IF GVL_HMI.rRobotManualSpeedPercent < REAL#0.1 THEN
	GVL_HMI.rRobotManualSpeedPercent := REAL#0.1;
ELSIF GVL_HMI.rRobotManualSpeedPercent > REAL#100.0 THEN
	GVL_HMI.rRobotManualSpeedPercent := REAL#100.0;
END_IF;
IF (GVL_HMI.lrRobotManualStep <> 0.1)
AND (GVL_HMI.lrRobotManualStep <> 1.0)
AND (GVL_HMI.lrRobotManualStep <> 10.0)
AND (GVL_HMI.lrRobotManualStep <> 100.0) THEN
	GVL_HMI.lrRobotManualStep := 1.0;
END_IF;

IF NOT xHmiConnectionAlive THEN
	FOR uiMachine := 1 TO 3 DO
		GVL_HMI.astAxisHmiCommand[uiMachine].xJogPositive := FALSE;
		GVL_HMI.astAxisHmiCommand[uiMachine].xJogNegative := FALSE;
		GVL_HMI.astAxisHmiCommand[uiMachine].xHome := FALSE;
		GVL_HMI.astAxisHmiCommand[uiMachine].xMoveAbsolute := FALSE;
		GVL_HMI.astAxisHmiCommand[uiMachine].xMoveRelative := FALSE;
	END_FOR;
	FOR uiMagazine := UINT#1 TO UINT#2 DO
		GVL_HMI.astMagazineCommand[uiMagazine].xStop := FALSE;
	END_FOR;
	GVL_HMI.xRobotManualExecute := FALSE;
END_IF;

// Глобальные команды ячейки поступают через единый интерфейс HMI.
GVL_CELL_CONTROL.xEnable := GVL_HMI.xCellEnable;
GVL_CELL_CONTROL.xDisable := GVL_HMI.xCellDisable;
GVL_CELL_CONTROL.xStart := GVL_HMI.xCellStart;
GVL_CELL_CONTROL.xStop := GVL_HMI.xCellStop;
// Необработанный общий импульс передаётся всем владельцам аварий.
// Каждый функциональный блок самостоятельно проверяет возможность сброса.
GVL_CELL_CONTROL.xReset := GVL_HMI.xCellReset;
// Режим хранит PLC. Новая транзакция применяется в RunSafety после чтения
// актуальных входов безопасности; PublishHmi не пишет в буфер запроса.
GVL_ALARM.Command.xResetWarnings := GVL_HMI.xAlarmResetWarnings;

// Режим инъекции ошибок включается отдельным переключателем страницы CELL_SETTINGS.
GVL_CELL_SETTINGS.xErrorSimulationEnabled := GVL_HMI.xErrorSimulationEnable
	AND (GVL_CELL_SETTINGS.eTestEnvironment <> E_CELL_TEST_ENVIRONMENT.NORMAL);

// Ползунок меняет только запрошенное значение. Отдельный FB применяет его к
// таймерам и Dynamic Limits безопасной транзакцией перед следующим тестом.
GVL_CELL_SETTINGS.xSimulationAccelerationChangeAllowed :=
	xHmiConnectionAlive
	AND NOT GVL_CELL_CONTROL.xGlobalError;

IF GVL_CELL_SETTINGS.xSimulationAccelerationChangeAllowed THEN
	GVL_CELL_SETTINGS.xSimulationAccelerationEnable := GVL_HMI.xSimulationAccelerationEnable;
	GVL_CELL_SETTINGS.uiSimulationTimeFactor := GVL_HMI.uiSimulationTimeFactor;
	IF GVL_CELL_SETTINGS.uiSimulationTimeFactor < UINT#1 THEN
		GVL_CELL_SETTINGS.uiSimulationTimeFactor := UINT#1;
	ELSIF GVL_CELL_SETTINGS.uiSimulationTimeFactor > UINT#100 THEN
		GVL_CELL_SETTINGS.uiSimulationTimeFactor := UINT#100;
	END_IF;
ELSE
	// При потере разрешения сохраняем последнее принятое требование.
	GVL_HMI.xSimulationAccelerationEnable := GVL_CELL_SETTINGS.xSimulationAccelerationActive;
	GVL_HMI.uiSimulationTimeFactor := GVL_CELL_SETTINGS.uiSimulationTimeFactor;
END_IF;

// Общие технологические TIMEOUT и допуски HOME принимаются только при полностью
// остановленной ячейке. Координатами HOME_SAFETY владеет редактор точек ниже.
GVL_CELL_SETTINGS.xCellSettingsChangeAllowed :=
	xHmiConnectionAlive
	AND NOT GVL_CELL_MANAGER.Status.xRunning
	AND NOT GVL_HMI.xModbusMode
	AND NOT GVL_CELL_CONTROL.xGlobalError
	AND NOT GVL_AXIS.arrAxis[1].Status.xMotionBusy
	AND NOT GVL_AXIS.arrAxis[2].Status.xMotionBusy
	AND NOT GVL_AXIS.arrAxis[3].Status.xMotionBusy
	AND NOT GVL_AXIS_GROUP.AxisGroup.Command.xMoveDirect
	AND NOT GVL_AXIS_GROUP.AxisGroup.Command.xMoveLinear
	AND NOT xPowerTransitionActive
	AND NOT SIMULATION_DYNAMICS.xBusy
	AND NOT GVL_ROBOT.Status.xBusy;

GVL_CELL_SETTINGS.xIoFilterSettingsChangeAllowed := xHmiConnectionAlive
	AND GVL_CELL_CONTROL.xManual
	AND NOT GVL_CELL_MANAGER.Status.xRunning
	AND NOT GVL_ROBOT.Status.xBusy AND NOT xMotionBusy
	AND NOT xPowerTransitionActive AND NOT SIMULATION_DYNAMICS.xBusy
	AND NOT GVL_MACHINE.Status[1].xBusy AND NOT GVL_MACHINE.Status[1].xProcessing
	AND NOT GVL_MACHINE.Status[2].xBusy AND NOT GVL_MACHINE.Status[2].xProcessing
	AND NOT GVL_MACHINE.Status[3].xBusy AND NOT GVL_MACHINE.Status[3].xProcessing
	AND NOT GVL_TWO_PALLET.astStatus[1].xBusy AND NOT GVL_TWO_PALLET.astStatus[2].xBusy
	AND NOT GVL_TWO_PALLET.astInput[1].xPowered AND NOT GVL_TWO_PALLET.astInput[2].xPowered;

// Independent requested value; publication cannot overwrite an incoming write.
xCellSettingRejected := FALSE;
udiCellSettingSnapshot := GVL_HMI.udiCellSettingCommandSeq;
IF (udiCellSettingSnapshot <> UDINT#0)
AND (udiCellSettingSnapshot <> GVL_HMI.udiCellSettingAckSeq) THEN
	GVL_HMI.uiCellSettingResult := UINT#3;
	IF NOT IsHmiCommandFresh(udiIssuedAtMs := GVL_HMI.udiCellSettingIssuedAtMs) THEN
		GVL_HMI.uiCellSettingResult := UINT#4; // Expired: never apply later
	ELSIF ((((GVL_HMI.uiCellSettingIndex = UINT#37) OR (GVL_HMI.uiCellSettingIndex = UINT#38) OR (GVL_HMI.uiCellSettingIndex = UINT#39))
		AND NOT GVL_CELL_SETTINGS.xIoFilterSettingsChangeAllowed)
		OR (((GVL_HMI.uiCellSettingIndex <> UINT#37) AND (GVL_HMI.uiCellSettingIndex <> UINT#38) AND (GVL_HMI.uiCellSettingIndex <> UINT#39))
			AND NOT GVL_CELL_SETTINGS.xCellSettingsChangeAllowed))
	OR (((GVL_HMI.uiCellSettingIndex = UINT#4)
		OR (GVL_HMI.uiCellSettingIndex = UINT#25)
		OR (GVL_HMI.uiCellSettingIndex = UINT#29))
		AND xPointCheckActive)
	OR ((GVL_HMI.uiCellSettingIndex = UINT#28) AND xMobileMotionLeaseActive) THEN
		GVL_HMI.uiCellSettingResult := UINT#2;
	ELSE
		CASE GVL_HMI.uiCellSettingIndex OF
			UINT#1:
				IF (GVL_HMI.lrCellSettingRequest >= 0.1) AND (GVL_HMI.lrCellSettingRequest <= 1000.0) THEN
					GVL_CELL_SETTINGS.lrSafetyHomeToleranceX := GVL_HMI.lrCellSettingRequest;
					GVL_HMI.uiCellSettingResult := UINT#1;
				END_IF;
			UINT#2:
				IF (GVL_HMI.lrCellSettingRequest >= 0.1) AND (GVL_HMI.lrCellSettingRequest <= 1000.0) THEN
					GVL_CELL_SETTINGS.lrSafetyHomeToleranceY := GVL_HMI.lrCellSettingRequest;
					GVL_HMI.uiCellSettingResult := UINT#1;
				END_IF;
			UINT#3:
				IF (GVL_HMI.lrCellSettingRequest >= 0.1) AND (GVL_HMI.lrCellSettingRequest <= 1000.0) THEN
					GVL_CELL_SETTINGS.lrSafetyHomeToleranceZ := GVL_HMI.lrCellSettingRequest;
					GVL_HMI.uiCellSettingResult := UINT#1;
				END_IF;
			UINT#4:
				IF (GVL_HMI.lrCellSettingRequest >= 0.1) AND (GVL_HMI.lrCellSettingRequest <= 100.0) THEN
					GVL_CELL_SETTINGS.rPointCheckSpeedPercent := LREAL_TO_REAL(GVL_HMI.lrCellSettingRequest);
					GVL_HMI.uiCellSettingResult := UINT#1;
				END_IF;
			UINT#5:
				IF (GVL_HMI.lrCellSettingRequest >= 1000.0) AND (GVL_HMI.lrCellSettingRequest <= 600000.0) THEN
					GVL_CELL_SETTINGS.stMachineTimeouts.tRobotMove := UDINT_TO_TIME(LREAL_TO_UDINT(GVL_HMI.lrCellSettingRequest));
					GVL_HMI.uiCellSettingResult := UINT#1;
				END_IF;
			UINT#6:
				IF (GVL_HMI.lrCellSettingRequest >= 1000.0) AND (GVL_HMI.lrCellSettingRequest <= 600000.0) THEN
					GVL_CELL_SETTINGS.stMachineTimeouts.tRobotAction := UDINT_TO_TIME(LREAL_TO_UDINT(GVL_HMI.lrCellSettingRequest));
					GVL_HMI.uiCellSettingResult := UINT#1;
				END_IF;
			UINT#7:
				IF (GVL_HMI.lrCellSettingRequest >= 1000.0) AND (GVL_HMI.lrCellSettingRequest <= 600000.0) THEN
					GVL_CELL_SETTINGS.stMachineTimeouts.tRobotRelease := UDINT_TO_TIME(LREAL_TO_UDINT(GVL_HMI.lrCellSettingRequest));
					GVL_HMI.uiCellSettingResult := UINT#1;
				END_IF;
			UINT#8:
				IF (GVL_HMI.lrCellSettingRequest >= 1000.0) AND (GVL_HMI.lrCellSettingRequest <= 600000.0) THEN
					GVL_CELL_SETTINGS.stMachineTimeouts.tDoorOpen := UDINT_TO_TIME(LREAL_TO_UDINT(GVL_HMI.lrCellSettingRequest));
					GVL_HMI.uiCellSettingResult := UINT#1;
				END_IF;
			UINT#9:
				IF (GVL_HMI.lrCellSettingRequest >= 1000.0) AND (GVL_HMI.lrCellSettingRequest <= 600000.0) THEN
					GVL_CELL_SETTINGS.stMachineTimeouts.tDoorClose := UDINT_TO_TIME(LREAL_TO_UDINT(GVL_HMI.lrCellSettingRequest));
					GVL_HMI.uiCellSettingResult := UINT#1;
				END_IF;
			UINT#10:
				IF (GVL_HMI.lrCellSettingRequest >= 1000.0) AND (GVL_HMI.lrCellSettingRequest <= 600000.0) THEN
					GVL_CELL_SETTINGS.stMachineTimeouts.tHatchUnlock := UDINT_TO_TIME(LREAL_TO_UDINT(GVL_HMI.lrCellSettingRequest));
					GVL_HMI.uiCellSettingResult := UINT#1;
				END_IF;
			UINT#11:
				IF (GVL_HMI.lrCellSettingRequest >= 1000.0) AND (GVL_HMI.lrCellSettingRequest <= 600000.0) THEN
					GVL_CELL_SETTINGS.stMachineTimeouts.tChuckOpen := UDINT_TO_TIME(LREAL_TO_UDINT(GVL_HMI.lrCellSettingRequest));
					GVL_HMI.uiCellSettingResult := UINT#1;
				END_IF;
			UINT#12:
				IF (GVL_HMI.lrCellSettingRequest >= 1000.0) AND (GVL_HMI.lrCellSettingRequest <= 600000.0) THEN
					GVL_CELL_SETTINGS.stMachineTimeouts.tChuckClose := UDINT_TO_TIME(LREAL_TO_UDINT(GVL_HMI.lrCellSettingRequest));
					GVL_HMI.uiCellSettingResult := UINT#1;
				END_IF;
			UINT#13:
				IF (GVL_HMI.lrCellSettingRequest >= 1000.0) AND (GVL_HMI.lrCellSettingRequest <= 600000.0) THEN
					GVL_CELL_SETTINGS.stMachineTimeouts.tCycleStart := UDINT_TO_TIME(LREAL_TO_UDINT(GVL_HMI.lrCellSettingRequest));
					GVL_HMI.uiCellSettingResult := UINT#1;
				END_IF;
			UINT#14:
				IF (GVL_HMI.lrCellSettingRequest >= 1000.0) AND (GVL_HMI.lrCellSettingRequest <= 600000.0) THEN
					GVL_CELL_SETTINGS.stAxisTimeouts.tPowerTimeout := UDINT_TO_TIME(LREAL_TO_UDINT(GVL_HMI.lrCellSettingRequest));
					GVL_HMI.uiCellSettingResult := UINT#1;
				END_IF;
			UINT#15:
				IF (GVL_HMI.lrCellSettingRequest >= 1000.0) AND (GVL_HMI.lrCellSettingRequest <= 600000.0) THEN
					GVL_CELL_SETTINGS.stAxisTimeouts.tResetTimeout := UDINT_TO_TIME(LREAL_TO_UDINT(GVL_HMI.lrCellSettingRequest));
					GVL_HMI.uiCellSettingResult := UINT#1;
				END_IF;
			UINT#16:
				IF (GVL_HMI.lrCellSettingRequest >= 1000.0) AND (GVL_HMI.lrCellSettingRequest <= 600000.0) THEN
					GVL_CELL_SETTINGS.stAxisTimeouts.tStopTimeout := UDINT_TO_TIME(LREAL_TO_UDINT(GVL_HMI.lrCellSettingRequest));
					GVL_HMI.uiCellSettingResult := UINT#1;
				END_IF;
			UINT#17:
				IF (GVL_HMI.lrCellSettingRequest >= 1000.0) AND (GVL_HMI.lrCellSettingRequest <= 600000.0) THEN
					GVL_CELL_SETTINGS.stAxisTimeouts.tHomeTimeout := UDINT_TO_TIME(LREAL_TO_UDINT(GVL_HMI.lrCellSettingRequest));
					GVL_HMI.uiCellSettingResult := UINT#1;
				END_IF;
			UINT#18:
				IF (GVL_HMI.lrCellSettingRequest >= 1000.0) AND (GVL_HMI.lrCellSettingRequest <= 600000.0) THEN
					GVL_CELL_SETTINGS.stAxisTimeouts.tMoveTimeout := UDINT_TO_TIME(LREAL_TO_UDINT(GVL_HMI.lrCellSettingRequest));
					GVL_HMI.uiCellSettingResult := UINT#1;
				END_IF;
			UINT#19:
				IF (GVL_HMI.lrCellSettingRequest >= 1000.0) AND (GVL_HMI.lrCellSettingRequest <= 600000.0) THEN
					GVL_CELL_SETTINGS.stAxisGroupTimeouts.tPowerTimeout := UDINT_TO_TIME(LREAL_TO_UDINT(GVL_HMI.lrCellSettingRequest));
					GVL_HMI.uiCellSettingResult := UINT#1;
				END_IF;
			UINT#20:
				IF (GVL_HMI.lrCellSettingRequest >= 1000.0) AND (GVL_HMI.lrCellSettingRequest <= 600000.0) THEN
					GVL_CELL_SETTINGS.stAxisGroupTimeouts.tGroupTimeout := UDINT_TO_TIME(LREAL_TO_UDINT(GVL_HMI.lrCellSettingRequest));
					GVL_HMI.uiCellSettingResult := UINT#1;
				END_IF;
			UINT#21:
				IF (GVL_HMI.lrCellSettingRequest >= 1000.0) AND (GVL_HMI.lrCellSettingRequest <= 600000.0) THEN
					GVL_CELL_SETTINGS.stAxisGroupTimeouts.tStopTimeout := UDINT_TO_TIME(LREAL_TO_UDINT(GVL_HMI.lrCellSettingRequest));
					GVL_HMI.uiCellSettingResult := UINT#1;
				END_IF;
			UINT#22:
				IF (GVL_HMI.lrCellSettingRequest >= 1000.0) AND (GVL_HMI.lrCellSettingRequest <= 600000.0) THEN
					GVL_CELL_SETTINGS.stAxisGroupTimeouts.tHaltTimeout := UDINT_TO_TIME(LREAL_TO_UDINT(GVL_HMI.lrCellSettingRequest));
					GVL_HMI.uiCellSettingResult := UINT#1;
				END_IF;
			UINT#23:
				IF (GVL_HMI.lrCellSettingRequest >= 1000.0) AND (GVL_HMI.lrCellSettingRequest <= 600000.0) THEN
					GVL_CELL_SETTINGS.stAxisGroupTimeouts.tHomeTimeout := UDINT_TO_TIME(LREAL_TO_UDINT(GVL_HMI.lrCellSettingRequest));
					GVL_HMI.uiCellSettingResult := UINT#1;
				END_IF;
			UINT#24:
				IF (GVL_HMI.lrCellSettingRequest >= 1000.0) AND (GVL_HMI.lrCellSettingRequest <= 600000.0) THEN
					GVL_CELL_SETTINGS.stAxisGroupTimeouts.tMoveTimeout := UDINT_TO_TIME(LREAL_TO_UDINT(GVL_HMI.lrCellSettingRequest));
					GVL_HMI.uiCellSettingResult := UINT#1;
				END_IF;
			UINT#25:
				IF (GVL_HMI.lrCellSettingRequest >= 500.0) AND (GVL_HMI.lrCellSettingRequest <= 60000.0) THEN
					GVL_CELL_SETTINGS.tPointCheckStartTimeout := UDINT_TO_TIME(LREAL_TO_UDINT(GVL_HMI.lrCellSettingRequest));
					GVL_HMI.uiCellSettingResult := UINT#1;
				END_IF;
			UINT#26:
				IF (GVL_HMI.lrCellSettingRequest >= 1000.0) AND (GVL_HMI.lrCellSettingRequest <= 600000.0) THEN
					GVL_CELL_SETTINGS.tSimulationDynamicsTimeout := UDINT_TO_TIME(LREAL_TO_UDINT(GVL_HMI.lrCellSettingRequest));
					GVL_HMI.uiCellSettingResult := UINT#1;
				END_IF;
			UINT#27:
				IF (GVL_HMI.lrCellSettingRequest >= 500.0) AND (GVL_HMI.lrCellSettingRequest <= 30000.0) THEN
					GVL_CELL_SETTINGS.tHmiWatchdogTimeout := UDINT_TO_TIME(LREAL_TO_UDINT(GVL_HMI.lrCellSettingRequest));
					GVL_HMI.uiCellSettingResult := UINT#1;
				END_IF;
			UINT#28:
				IF (GVL_HMI.lrCellSettingRequest >= 500.0) AND (GVL_HMI.lrCellSettingRequest <= 30000.0) THEN
					GVL_CELL_SETTINGS.tMobileMotionWatchdogTimeout := UDINT_TO_TIME(LREAL_TO_UDINT(GVL_HMI.lrCellSettingRequest));
					GVL_HMI.uiCellSettingResult := UINT#1;
				END_IF;
			UINT#29:
				IF (GVL_HMI.lrCellSettingRequest >= 500.0) AND (GVL_HMI.lrCellSettingRequest <= 30000.0) THEN
					GVL_CELL_SETTINGS.tPointCheckWatchdogTimeout := UDINT_TO_TIME(LREAL_TO_UDINT(GVL_HMI.lrCellSettingRequest));
					GVL_HMI.uiCellSettingResult := UINT#1;
				END_IF;
			UINT#30:
				IF (GVL_HMI.lrCellSettingRequest >= 1000.0) AND (GVL_HMI.lrCellSettingRequest <= 30000.0) THEN
					GVL_CELL_SETTINGS.tHmiCommandFreshnessTimeout := UDINT_TO_TIME(LREAL_TO_UDINT(GVL_HMI.lrCellSettingRequest));
					GVL_HMI.uiCellSettingResult := UINT#1;
				END_IF;
			UINT#31:
				IF (GVL_HMI.lrCellSettingRequest >= 100.0) AND (GVL_HMI.lrCellSettingRequest <= 10000.0) THEN
					GVL_CELL_SETTINGS.stAxisTimeouts.tPowerFeedbackLossTimeout := UDINT_TO_TIME(LREAL_TO_UDINT(GVL_HMI.lrCellSettingRequest));
					GVL_HMI.uiCellSettingResult := UINT#1;
				END_IF;
			UINT#32:
				IF (GVL_HMI.lrCellSettingRequest >= 1.0) AND (GVL_HMI.lrCellSettingRequest <= 100.0) THEN
					GVL_CELL_SETTINGS.rRobotAccelerationPercent := LREAL_TO_REAL(GVL_HMI.lrCellSettingRequest);
					GVL_HMI.uiCellSettingResult := UINT#1;
				END_IF;
			UINT#33:
				IF (GVL_HMI.lrCellSettingRequest >= 1.0) AND (GVL_HMI.lrCellSettingRequest <= 100.0) THEN
					GVL_CELL_SETTINGS.rRobotDecelerationPercent := LREAL_TO_REAL(GVL_HMI.lrCellSettingRequest);
					GVL_HMI.uiCellSettingResult := UINT#1;
				END_IF;
			UINT#34:
				IF (GVL_HMI.lrCellSettingRequest >= 1.0) AND (GVL_HMI.lrCellSettingRequest <= 100.0) THEN
					GVL_CELL_SETTINGS.rRobotJerkPercent := LREAL_TO_REAL(GVL_HMI.lrCellSettingRequest);
					GVL_HMI.uiCellSettingResult := UINT#1;
				END_IF;
			UINT#35:
				IF (GVL_HMI.lrCellSettingRequest >= 1.0) AND (GVL_HMI.lrCellSettingRequest <= 100000.0) THEN
					GVL_CELL_SETTINGS.lrRobotHaltDeceleration := GVL_HMI.lrCellSettingRequest;
					GVL_HMI.uiCellSettingResult := UINT#1;
				END_IF;
			UINT#36:
				IF (GVL_HMI.lrCellSettingRequest >= 1.0) AND (GVL_HMI.lrCellSettingRequest <= 1000000.0) THEN
					GVL_CELL_SETTINGS.lrRobotHaltJerk := GVL_HMI.lrCellSettingRequest;
					GVL_HMI.uiCellSettingResult := UINT#1;
				END_IF;
			UINT#37:
				IF (GVL_HMI.lrCellSettingRequest >= 0.0) AND (GVL_HMI.lrCellSettingRequest <= 5000.0) THEN
					GVL_CELL_SETTINGS.tInputFilterRise := UDINT_TO_TIME(LREAL_TO_UDINT(GVL_HMI.lrCellSettingRequest));
					GVL_HMI.uiCellSettingResult := UINT#1;
				END_IF;
			UINT#38:
				IF (GVL_HMI.lrCellSettingRequest >= 0.0) AND (GVL_HMI.lrCellSettingRequest <= 5000.0) THEN
					GVL_CELL_SETTINGS.tInputFilterFall := UDINT_TO_TIME(LREAL_TO_UDINT(GVL_HMI.lrCellSettingRequest));
					GVL_HMI.uiCellSettingResult := UINT#1;
				END_IF;
			UINT#39:
				IF (GVL_HMI.lrCellSettingRequest >= 0.0) AND (GVL_HMI.lrCellSettingRequest <= 60000.0) THEN
					GVL_CELL_SETTINGS.tAlarmHornDuration := UDINT_TO_TIME(LREAL_TO_UDINT(GVL_HMI.lrCellSettingRequest));
					GVL_HMI.uiCellSettingResult := UINT#1;
				END_IF;
		END_CASE;
	END_IF;
	xCellSettingRejected := GVL_HMI.uiCellSettingResult <> UINT#1;
END_IF;

// =============================================================================
// Транзакционный редактор 14 фиксированных инженерных точек
// =============================================================================
xPointEditorAllHomed := GVL_AXIS.arrAxis[1].Status.xHomed
	AND GVL_AXIS.arrAxis[2].Status.xHomed
	AND GVL_AXIS.arrAxis[3].Status.xHomed;
xPointEditorBaseAllowed := xHmiConnectionAlive
	AND NOT xPointCheckActive
	AND GVL_CELL_CONTROL.xManual
	AND NOT GVL_HMI.xModbusMode
	AND NOT GVL_CELL_MANAGER.Status.xRunning
	AND NOT GVL_CELL_CONTROL.xGlobalError
	AND NOT GVL_ROBOT.Status.xBusy
	AND NOT xMotionBusy
	AND NOT xDriveError
	AND NOT GVL_MOTION_MANAGER.stMotionManager.Status.xError
	AND xPointEditorAllHomed
	AND GVL_AXIS_GROUP.AxisGroup.Status.xPositionValid;
GVL_HMI.xPointEditorCaptureAllowed := xPointEditorBaseAllowed;
GVL_HMI.xPointEditorSaveAllowed := xPointEditorBaseAllowed
	AND GVL_POINT_MANAGER.PointManager.Diag.xXLimitValid
	AND GVL_POINT_MANAGER.PointManager.Diag.xYLimitValid
	AND GVL_POINT_MANAGER.PointManager.Diag.xZLimitValid;

IF (GVL_HMI.udiPointEditorCommandSeq <> UDINT#0)
AND (GVL_HMI.udiPointEditorCommandSeq <> udiLastPointEditorCommandSeq) THEN
	udiLastPointEditorCommandSeq := GVL_HMI.udiPointEditorCommandSeq;
	GVL_HMI.uiPointEditorResult := UINT#2;
	GVL_HMI.uiPointEditorRejectReason := UINT#0;
	xPointEditorRequestValid := FALSE;
	xPointEditorMagazinePoint := FALSE;
	uiPointEditorGeometryStation := UINT#0;
	ePointEditorName := E_POINT_NAME.NONE;
	uiPointStorageIndex := UINT#0;

	CASE GVL_HMI.uiPointEditorIndex OF
		UINT#1: ePointEditorName := E_POINT_NAME.MACHINE_1_ABOVE; uiPointStorageIndex := UINT#1;
		UINT#2: ePointEditorName := E_POINT_NAME.MACHINE_1_CHUCK_APROACH; uiPointStorageIndex := UINT#3;
		UINT#3: ePointEditorName := E_POINT_NAME.MACHINE_1_CHUCK_POSITION; uiPointStorageIndex := UINT#4;
		UINT#4: ePointEditorName := E_POINT_NAME.MACHINE_2_ABOVE; uiPointStorageIndex := UINT#5;
		UINT#5: ePointEditorName := E_POINT_NAME.MACHINE_2_CHUCK_APROACH; uiPointStorageIndex := UINT#7;
		UINT#6: ePointEditorName := E_POINT_NAME.MACHINE_2_CHUCK_POSITION; uiPointStorageIndex := UINT#8;
		UINT#7: ePointEditorName := E_POINT_NAME.MACHINE_3_ABOVE; uiPointStorageIndex := UINT#9;
		UINT#8: ePointEditorName := E_POINT_NAME.MACHINE_3_CHUCK_APROACH; uiPointStorageIndex := UINT#11;
		UINT#9: ePointEditorName := E_POINT_NAME.MACHINE_3_CHUCK_POSITION; uiPointStorageIndex := UINT#12;
		UINT#10: ePointEditorName := E_POINT_NAME.HOME_SAFETY; uiPointStorageIndex := UINT#13;
		UINT#11: ePointEditorName := E_POINT_NAME.MAGAZINE_1_DETAIL; uiPointStorageIndex := UINT#14;
		UINT#12: ePointEditorName := E_POINT_NAME.MAGAZINE_2_DETAIL; uiPointStorageIndex := UINT#15;
		UINT#13: ePointEditorName := E_POINT_NAME.GEOMETRY_1_PLACE; uiPointEditorGeometryStation := UINT#1;
		UINT#14: ePointEditorName := E_POINT_NAME.GEOMETRY_2_PLACE; uiPointEditorGeometryStation := UINT#2;
	END_CASE;
	xPointEditorRequestValid := (ePointEditorName <> E_POINT_NAME.NONE)
		AND ((uiPointStorageIndex <> UINT#0) OR (uiPointEditorGeometryStation <> UINT#0));
	xPointEditorMagazinePoint := (ePointEditorName = E_POINT_NAME.MAGAZINE_1_DETAIL)
		OR (ePointEditorName = E_POINT_NAME.MAGAZINE_2_DETAIL);
	xPointEditorGeometrySave := (GVL_HMI.uiPointEditorCommand = UINT#2)
		AND (uiPointEditorGeometryStation <> UINT#0);

	IF (GVL_HMI.uiPointEditorCommand <> UINT#1)
	AND (GVL_HMI.uiPointEditorCommand <> UINT#2)
	AND (GVL_HMI.uiPointEditorCommand <> UINT#3) THEN
		GVL_HMI.uiPointEditorRejectReason := UINT#1; // Неизвестная команда
	ELSIF NOT xPointEditorRequestValid THEN
		GVL_HMI.uiPointEditorRejectReason := UINT#2; // Неверный индекс точки
	ELSIF NOT xHmiConnectionAlive THEN
		GVL_HMI.uiPointEditorRejectReason := UINT#3; // HMI offline
	ELSIF xPointEditorGeometrySave THEN
		// SAVE только изменяет данные. Режим, Home, движение, ошибки и состояние
		// ГК не блокируют запись. CAPTURE/CHECK сохраняют прежние допуски.
		IF GVL_HMI.xModbusMode
		OR (GVL_CELL_SETTINGS.eTestEnvironment = E_CELL_TEST_ENVIRONMENT.SC500_BENCH) THEN
			GVL_HMI.uiPointEditorRejectReason := UINT#5;
		ELSIF NOT GVL_POINT_MANAGER.PointManager.Diag.xXLimitValid
		OR NOT GVL_POINT_MANAGER.PointManager.Diag.xYLimitValid
		OR NOT GVL_POINT_MANAGER.PointManager.Diag.xZLimitValid THEN
			GVL_HMI.uiPointEditorRejectReason := UINT#13;
		END_IF;
	ELSIF NOT GVL_CELL_CONTROL.xManual THEN
		GVL_HMI.uiPointEditorRejectReason := UINT#4; // Требуется ручной режим
	ELSIF GVL_HMI.xModbusMode THEN
		GVL_HMI.uiPointEditorRejectReason := UINT#5; // Требуется SoftMotion
	ELSIF GVL_CELL_MANAGER.Status.xRunning THEN
		GVL_HMI.uiPointEditorRejectReason := UINT#6; // Автоматический цикл выполняется
	ELSIF GVL_CELL_CONTROL.xGlobalError THEN
		GVL_HMI.uiPointEditorRejectReason := UINT#7; // Глобальная ошибка
	ELSIF GVL_ROBOT.Status.xBusy OR xPointCheckActive THEN
		GVL_HMI.uiPointEditorRejectReason := UINT#8; // Робот занят
	ELSIF xMotionBusy THEN
		GVL_HMI.uiPointEditorRejectReason := UINT#9; // Motion занят
	ELSIF xDriveError OR GVL_MOTION_MANAGER.stMotionManager.Status.xError THEN
		GVL_HMI.uiPointEditorRejectReason := UINT#10; // Ошибка оси или группы
	ELSIF NOT xPointEditorAllHomed THEN
		GVL_HMI.uiPointEditorRejectReason := UINT#11; // Не выполнен Home
	ELSIF NOT GVL_AXIS_GROUP.AxisGroup.Status.xPositionValid THEN
		GVL_HMI.uiPointEditorRejectReason := UINT#12; // Недостоверные координаты
	ELSIF (GVL_HMI.uiPointEditorCommand = UINT#2)
	AND (NOT GVL_POINT_MANAGER.PointManager.Diag.xXLimitValid
		OR NOT GVL_POINT_MANAGER.PointManager.Diag.xYLimitValid
		OR NOT GVL_POINT_MANAGER.PointManager.Diag.xZLimitValid) THEN
		GVL_HMI.uiPointEditorRejectReason := UINT#13; // Software limits недоступны
	END_IF;

	IF GVL_HMI.uiPointEditorRejectReason = UINT#0 THEN
		IF GVL_HMI.uiPointEditorCommand = UINT#1 THEN
			// CAPTURE возвращает согласованный снимок одного PLC-цикла и не пишет Persistent.
			GVL_HMI.stPointEditorResultPoint.Name := '';
			GVL_HMI.stPointEditorResultPoint.X := GVL_AXIS_GROUP.AxisGroup.Status.ActualX;
			GVL_HMI.stPointEditorResultPoint.Y := GVL_AXIS_GROUP.AxisGroup.Status.ActualY;
			GVL_HMI.stPointEditorResultPoint.Z := GVL_AXIS_GROUP.AxisGroup.Status.ActualZ;
			GVL_HMI.stPointEditorResultPoint.MagazineSafeZ :=
				GVL_HMI.lrPointEditorDraftMagazineSafeZ;
			GVL_HMI.stPointEditorResultPoint.MagazineChangeZ :=
				GVL_HMI.lrPointEditorDraftMagazineChangeZ;
			GVL_HMI.stPointEditorResultPoint.SpeedFactor :=
				GVL_HMI.lrPointEditorDraftSpeedFactor;
			GVL_HMI.stPointEditorResultPoint.xConfigured := FALSE;
			GVL_HMI.uiPointEditorResult := UINT#1;
		ELSIF GVL_HMI.uiPointEditorCommand = UINT#3 THEN
			// CHECK никогда не сохраняет черновик. Сравнение защищает подтверждение
			// на телефоне от изменения точки другим редактором до запуска.
			IF NOT GVL_POINT.Points[ePointEditorName].xConfigured THEN
				GVL_HMI.uiPointEditorRejectReason := UINT#16;
			ELSIF (GVL_POINT.Points[ePointEditorName].X <> GVL_HMI.alrPointEditorDraftXYZ[1])
			OR (GVL_POINT.Points[ePointEditorName].Y <> GVL_HMI.alrPointEditorDraftXYZ[2])
			OR (GVL_POINT.Points[ePointEditorName].Z <> GVL_HMI.alrPointEditorDraftXYZ[3])
			OR (GVL_POINT.Points[ePointEditorName].SpeedFactor <> GVL_HMI.lrPointEditorDraftSpeedFactor)
			OR ((xPointEditorMagazinePoint OR (uiPointEditorGeometryStation <> UINT#0))
				AND ((GVL_POINT.Points[ePointEditorName].MagazineSafeZ <>
					GVL_HMI.lrPointEditorDraftMagazineSafeZ)
				OR (GVL_POINT.Points[ePointEditorName].MagazineChangeZ <>
					GVL_HMI.lrPointEditorDraftMagazineChangeZ))) THEN
				GVL_HMI.uiPointEditorRejectReason := UINT#21;
			ELSE
				xPointCheckRequest := TRUE; // Финальное разрешение после RunMotion/RunCellControl
			END_IF;
		ELSE
			xPointEditorDraftValid :=
				(GVL_HMI.alrPointEditorDraftXYZ[1] >= alrRobotSoftwareMinPosition[1])
				AND (GVL_HMI.alrPointEditorDraftXYZ[1] <= alrRobotSoftwareMaxPosition[1])
				AND (GVL_HMI.alrPointEditorDraftXYZ[2] >= alrRobotSoftwareMinPosition[2])
				AND (GVL_HMI.alrPointEditorDraftXYZ[2] <= alrRobotSoftwareMaxPosition[2])
				AND (GVL_HMI.alrPointEditorDraftXYZ[3] >= alrRobotSoftwareMinPosition[3])
				AND (GVL_HMI.alrPointEditorDraftXYZ[3] <= alrRobotSoftwareMaxPosition[3]);
			IF NOT xPointEditorDraftValid THEN
				GVL_HMI.uiPointEditorRejectReason := UINT#14; // XYZ вне software limits
			ELSIF NOT (((GVL_HMI.lrPointEditorDraftSpeedFactor > 0.1)
				OR ((uiPointEditorGeometryStation <> UINT#0) AND (GVL_HMI.lrPointEditorDraftSpeedFactor >= 0.1)))
			AND (GVL_HMI.lrPointEditorDraftSpeedFactor <= 1.0)) THEN
				GVL_HMI.uiPointEditorRejectReason := UINT#15; // Недопустимая скорость
			ELSIF xPointEditorMagazinePoint
			AND ((GVL_HMI.lrPointEditorDraftMagazineSafeZ < -LREAL#10000.0)
				OR (GVL_HMI.lrPointEditorDraftMagazineSafeZ > LREAL#10000.0)
				OR (GVL_HMI.lrPointEditorDraftMagazineChangeZ < -LREAL#10000.0)
				OR (GVL_HMI.lrPointEditorDraftMagazineChangeZ > LREAL#10000.0)) THEN
				GVL_HMI.uiPointEditorRejectReason := UINT#22; // Смещения магазина вне диапазона
			ELSIF (uiPointEditorGeometryStation <> UINT#0)
			AND NOT ((GVL_HMI.lrPointEditorDraftMagazineSafeZ < LREAL#0.0)
				AND (GVL_HMI.lrPointEditorDraftMagazineSafeZ >= -LREAL#10000.0)
				AND ((GVL_HMI.alrPointEditorDraftXYZ[3] + GVL_HMI.lrPointEditorDraftMagazineSafeZ) >= alrRobotSoftwareMinPosition[3])
				AND ((GVL_HMI.alrPointEditorDraftXYZ[3] + GVL_HMI.lrPointEditorDraftMagazineSafeZ) <= alrRobotSoftwareMaxPosition[3])) THEN
				GVL_HMI.uiPointEditorRejectReason := UINT#22; // SAFE_Z ГК должен поднимать робот в пределах оси
			ELSIF uiPointEditorGeometryStation <> UINT#0 THEN
				// Единственный владелец базы ГК: действующая конфигурация NORMAL/SIMULATION.
				stGeometryConfig.lrX := GVL_HMI.alrPointEditorDraftXYZ[1];
				stGeometryConfig.lrY := GVL_HMI.alrPointEditorDraftXYZ[2];
				stGeometryConfig.lrZ := GVL_HMI.alrPointEditorDraftXYZ[3];
				stGeometryConfig.lrSafeZ := GVL_HMI.lrPointEditorDraftMagazineSafeZ;
				stGeometryConfig.lrChangeZ := stGeometryConfig.lrSafeZ; // Совместимый legacy-канал, отдельного CHANGE нет
				stGeometryConfig.lrSpeedFactor := GVL_HMI.lrPointEditorDraftSpeedFactor;
				stGeometryConfig.xConfigured := TRUE;
				IF GVL_CELL_SETTINGS.eTestEnvironment = E_CELL_TEST_ENVIRONMENT.NORMAL THEN
					GVL_GEOMETRY_CONTROL.astConfig[uiPointEditorGeometryStation] := stGeometryConfig;
				ELSE
					GVL_GEOMETRY_CONTROL.astSimulationConfig[uiPointEditorGeometryStation] := stGeometryConfig;
				END_IF;
				GVL_GEOMETRY_CONTROL.astActiveConfig[uiPointEditorGeometryStation] := stGeometryConfig;
				GVL_HMI.stPointEditorResultPoint.Name := '';
				GVL_HMI.stPointEditorResultPoint.X := stGeometryConfig.lrX;
				GVL_HMI.stPointEditorResultPoint.Y := stGeometryConfig.lrY;
				GVL_HMI.stPointEditorResultPoint.Z := stGeometryConfig.lrZ;
				GVL_HMI.stPointEditorResultPoint.MagazineSafeZ := stGeometryConfig.lrSafeZ;
				GVL_HMI.stPointEditorResultPoint.MagazineChangeZ := LREAL#0.0;
				GVL_HMI.stPointEditorResultPoint.SpeedFactor := stGeometryConfig.lrSpeedFactor;
				GVL_HMI.stPointEditorResultPoint.xConfigured := TRUE;
				GVL_HMI.uiPointEditorResult := UINT#1;
			ELSE
				GVL_POINT.astRetainPoints[uiPointStorageIndex].Name := '';
				GVL_POINT.astRetainPoints[uiPointStorageIndex].X :=
					GVL_HMI.alrPointEditorDraftXYZ[1];
				GVL_POINT.astRetainPoints[uiPointStorageIndex].Y :=
					GVL_HMI.alrPointEditorDraftXYZ[2];
				GVL_POINT.astRetainPoints[uiPointStorageIndex].Z :=
					GVL_HMI.alrPointEditorDraftXYZ[3];
				IF xPointEditorMagazinePoint THEN
					GVL_POINT.astRetainPoints[uiPointStorageIndex].MagazineSafeZ :=
						GVL_HMI.lrPointEditorDraftMagazineSafeZ;
					GVL_POINT.astRetainPoints[uiPointStorageIndex].MagazineChangeZ :=
						GVL_HMI.lrPointEditorDraftMagazineChangeZ;
				ELSE
					GVL_POINT.astRetainPoints[uiPointStorageIndex].MagazineSafeZ := LREAL#0.0;
					GVL_POINT.astRetainPoints[uiPointStorageIndex].MagazineChangeZ := LREAL#0.0;
				END_IF;
				GVL_POINT.astRetainPoints[uiPointStorageIndex].SpeedFactor :=
					GVL_HMI.lrPointEditorDraftSpeedFactor;
				GVL_POINT.astRetainPoints[uiPointStorageIndex].xConfigured :=
					NOT xPointEditorMagazinePoint
					OR ((GVL_HMI.lrPointEditorDraftMagazineSafeZ <> LREAL#0.0)
						AND (GVL_HMI.lrPointEditorDraftMagazineChangeZ <> LREAL#0.0));
				GVL_POINT.Points[ePointEditorName] :=
					GVL_POINT.astRetainPoints[uiPointStorageIndex];
				GVL_HMI.stPointEditorResultPoint := GVL_POINT.Points[ePointEditorName];
				GVL_HMI.uiPointEditorResult := UINT#1;
			END_IF;
		END_IF;
	END_IF;

	IF (GVL_HMI.uiPointEditorResult <> UINT#1) AND NOT xPointCheckRequest THEN
		IF GVL_HMI.uiPointEditorCommand = UINT#3 THEN
			uiRobotInterfaceWarningCode := WRN_POINT_CHECK_REJECTED;
		ELSE
			uiRobotInterfaceWarningCode := WRN_POINT_EDIT_REJECTED;
		END_IF;
	END_IF;
	// Ack подтверждает обработку конкретной транзакции даже при отказе.
	IF NOT xPointCheckRequest THEN
		GVL_HMI.udiPointEditorAckSeq := GVL_HMI.udiPointEditorCommandSeq;
	END_IF;
END_IF;

// Плоский OPC UA-интерфейс HMI преобразуется в типизированные запросы FB.
FOR uiMachine := 1 TO 3 DO
	astMachineFaultRequest[uiMachine].xEnabled := GVL_CELL_SETTINGS.xErrorSimulationEnabled;
	astMachineFaultRequest[uiMachine].xReset := GVL_HMI.axMachineSimReset[uiMachine];
	astMachineFaultRequest[uiMachine].xMachineAlarm := GVL_HMI.axMachineSimAlarm[uiMachine];
	astMachineFaultRequest[uiMachine].xDoorFault := GVL_HMI.axMachineSimDoorFault[uiMachine];
	astMachineFaultRequest[uiMachine].xChuckFault := GVL_HMI.axMachineSimChuckFault[uiMachine];
	astMachineFaultRequest[uiMachine].xTimeoutRobotMove := GVL_HMI.axMachineTimeoutRobotMove[uiMachine];
	astMachineFaultRequest[uiMachine].xTimeoutRobotAction := GVL_HMI.axMachineTimeoutRobotAction[uiMachine];
	astMachineFaultRequest[uiMachine].xTimeoutRobotRelease := GVL_HMI.axMachineTimeoutRobotRelease[uiMachine];
	astMachineFaultRequest[uiMachine].xTimeoutDoorOpen := GVL_HMI.axMachineTimeoutDoorOpen[uiMachine];
	astMachineFaultRequest[uiMachine].xTimeoutDoorClose := GVL_HMI.axMachineTimeoutDoorClose[uiMachine];
	astMachineFaultRequest[uiMachine].xTimeoutHatchUnlock := GVL_HMI.axMachineTimeoutHatchUnlock[uiMachine];
	astMachineFaultRequest[uiMachine].xTimeoutChuckOpen := GVL_HMI.axMachineTimeoutChuckOpen[uiMachine];
	astMachineFaultRequest[uiMachine].xTimeoutChuckClose := GVL_HMI.axMachineTimeoutChuckClose[uiMachine];
	astMachineFaultRequest[uiMachine].xTimeoutCycleStart := GVL_HMI.axMachineTimeoutCycleStart[uiMachine];

	astAxisFaultRequest[uiMachine].xEnabled := GVL_CELL_SETTINGS.xErrorSimulationEnabled;
	astAxisFaultRequest[uiMachine].xJogConflict := GVL_HMI.axSimAxisJogConflict[uiMachine];
END_FOR;

stAxisGroupFaultRequest.xEnabled := GVL_CELL_SETTINGS.xErrorSimulationEnabled;
stAxisGroupFaultRequest.xExecute := GVL_HMI.xSimAxisGroupError;

stRobotFaultRequest.xEnabled := GVL_CELL_SETTINGS.xErrorSimulationEnabled;
stRobotFaultRequest.xWrongAction := GVL_HMI.xSimRobotWrongAction;
stRobotFaultRequest.stGripper.xEnabled := GVL_CELL_SETTINGS.xErrorSimulationEnabled;
stRobotFaultRequest.stGripper.xGripper1Fault := GVL_HMI.xSimGripper1Fault;
stRobotFaultRequest.stGripper.xGripper2Fault := GVL_HMI.xSimGripper2Fault;
stRobotFaultRequest.stGripper.xRotationFault := GVL_HMI.xSimGripperRotationFault;
stRobotFaultRequest.stGripper.xGlobalFault := GVL_HMI.xSimGripperGlobalFault;

stRobotFaultRequest.stPoint.xEnabled := GVL_CELL_SETTINGS.xErrorSimulationEnabled;
stRobotFaultRequest.stPoint.xXOutOfLimit := GVL_HMI.xSimPointXOutOfLimit;
stRobotFaultRequest.stPoint.xYOutOfLimit := GVL_HMI.xSimPointYOutOfLimit;
stRobotFaultRequest.stPoint.xZOutOfLimit := GVL_HMI.xSimPointZOutOfLimit;
stRobotFaultRequest.stPoint.xInvalidVelocity := GVL_HMI.xSimPointInvalidVelocity;

IF NOT GVL_CELL_SETTINGS.xErrorSimulationEnabled THEN
	adwTestMagazineFaultMask[1] := DWORD#0;
	adwTestMagazineFaultMask[2] := DWORD#0;
END_IF;
astMagazineFaultRequest[1].xEnabled := GVL_CELL_SETTINGS.xErrorSimulationEnabled;
astMagazineFaultRequest[1].xWrongOperation := GVL_HMI.xSimMagazineWrongOperation
	OR ((adwTestMagazineFaultMask[1] AND DWORD#16#0000_0001) <> DWORD#0);
astMagazineFaultRequest[1].xNoBlank := GVL_HMI.xSimMagazineNoBlank
	OR ((adwTestMagazineFaultMask[1] AND DWORD#16#0000_0002) <> DWORD#0);
astMagazineFaultRequest[1].xNoFreeSlot := GVL_HMI.xSimMagazineNoFreeSlot
	OR ((adwTestMagazineFaultMask[1] AND DWORD#16#0000_0004) <> DWORD#0);
astMagazineFaultRequest[1].xInvalidSlot := GVL_HMI.xSimMagazineInvalidSlot
	OR ((adwTestMagazineFaultMask[1] AND DWORD#16#0000_0008) <> DWORD#0);
astMagazineFaultRequest[1].xSlotContent := GVL_HMI.xSimMagazineSlotContent
	OR ((adwTestMagazineFaultMask[1] AND DWORD#16#0000_0010) <> DWORD#0);
astMagazineFaultRequest[1].xGeometry := GVL_HMI.xSimMagazineGeometry
	OR ((adwTestMagazineFaultMask[1] AND DWORD#16#0000_0020) <> DWORD#0);
astMagazineFaultRequest[2].xEnabled := GVL_CELL_SETTINGS.xErrorSimulationEnabled
	AND (adwTestMagazineFaultMask[2] <> DWORD#0);
astMagazineFaultRequest[2].xWrongOperation :=
	(adwTestMagazineFaultMask[2] AND DWORD#16#0000_0001) <> DWORD#0;
astMagazineFaultRequest[2].xNoBlank :=
	(adwTestMagazineFaultMask[2] AND DWORD#16#0000_0002) <> DWORD#0;
astMagazineFaultRequest[2].xNoFreeSlot :=
	(adwTestMagazineFaultMask[2] AND DWORD#16#0000_0004) <> DWORD#0;
astMagazineFaultRequest[2].xInvalidSlot :=
	(adwTestMagazineFaultMask[2] AND DWORD#16#0000_0008) <> DWORD#0;
astMagazineFaultRequest[2].xSlotContent :=
	(adwTestMagazineFaultMask[2] AND DWORD#16#0000_0010) <> DWORD#0;
astMagazineFaultRequest[2].xGeometry :=
	(adwTestMagazineFaultMask[2] AND DWORD#16#0000_0020) <> DWORD#0;

stCellFaultRequest.xEnabled := GVL_CELL_SETTINGS.xErrorSimulationEnabled;
stCellFaultRequest.xBothGrippers := GVL_HMI.xSimCellBothGrippers;

stSafetyFaultRequest.xEnabled := GVL_CELL_SETTINGS.xErrorSimulationEnabled;
FOR uiMachine := UINT#1 TO UINT#4 DO
	stSafetyFaultRequest.axEmergencyStopStation[uiMachine] :=
		GVL_HMI.axSimSafetyEmergencyStopStation[uiMachine];
	stSafetyFaultRequest.axDoorUnlocked[uiMachine] :=
		GVL_HMI.axSimSafetyDoorUnlocked[uiMachine];
END_FOR;
FOR uiMachine := UINT#1 TO UINT#2 DO
	stSafetyFaultRequest.axEmergencyStopCabinet[uiMachine] :=
		GVL_HMI.axSimSafetyEmergencyStopCabinet[uiMachine];
END_FOR;
stSafetyFaultRequest.xEmergencyStopMpg := GVL_HMI.xSimSafetyEmergencyStopMpg;
stSafetyFaultRequest.xPhaseRelayFault := GVL_HMI.xSimSafetyPhaseRelayFault;
stSafetyFaultRequest.xPressureRelayFault := GVL_HMI.xSimSafetyPressureRelayFault;
stSafetyFaultRequest.xSafetyRelayFault := GVL_HMI.xSimSafetyRelayFault;
END_METHOD

METHOD PRIVATE ResetIoEmergencyStop
// Сырые аппаратные сигналы используются для снятия программного останова.
// Прямое ручное I/O этим условием не блокируется.
xIoRawSafetyOk := GVL_PHYSICAL_IO.xMappingVerified
    AND GVL_PHYSICAL_IO.xDiEmergencyStopStation1Ok
    AND GVL_PHYSICAL_IO.xDiEmergencyStopStation2Ok
    AND GVL_PHYSICAL_IO.xDiEmergencyStopStation3Ok
    AND GVL_PHYSICAL_IO.xDiEmergencyStopStation4Ok
    AND GVL_PHYSICAL_IO.xDiEmergencyStopCabinet1Ok
    AND GVL_PHYSICAL_IO.xDiEmergencyStopCabinet2Ok
    AND GVL_PHYSICAL_IO.xDiEmergencyStopMpgOk
    AND GVL_PHYSICAL_IO.xDiSafetyRelayOkInput
    AND GVL_PHYSICAL_IO.xDiPhaseRelayOkInput
    AND GVL_PHYSICAL_IO.xDiPressureRelayOkInput;
// Снять программный останов можно только после останова. Снятие не запускает механизм.
GVL_HMI.xIoEmergencyResetAllowed := GVL_HMI.xIoEmergencyStopActive
    AND GVL_CELL_CONTROL.xManual AND NOT xIoBusy AND xHmiConnectionAlive
    AND CELL_SAFETY.Status.xReady
    AND ((GVL_CELL_SETTINGS.eTestEnvironment <> E_CELL_TEST_ENVIRONMENT.NORMAL) OR xIoRawSafetyOk);
IF GVL_HMI.xIoEmergencyStopActive THEN
    GVL_CELL_CONTROL.xStart := FALSE;
    GVL_CELL_CONTROL.xEnable := FALSE;
    GVL_CELL_CONTROL.xManual := TRUE;
    xRobotHmiPermit := FALSE;
END_IF;
IF xIoEmergencyResetRequested THEN
    GVL_HMI.uiIoEmergencyResult := UINT#3;
    IF NOT IsHmiCommandFresh(udiIssuedAtMs := GVL_HMI.udiIoEmergencyIssuedAtMs) THEN
        GVL_HMI.uiIoEmergencyResult := UINT#4;
    ELSIF GVL_HMI.uiIoEmergencyAction = UINT#2 THEN
        IF GVL_HMI.xIoEmergencyResetAllowed THEN
            GVL_HMI.xIoEmergencyStopActive := FALSE;
            GVL_HMI.uiIoEmergencyResult := UINT#1;
        ELSE GVL_HMI.uiIoEmergencyResult := UINT#2;
        END_IF;
    END_IF;
    xIoEmergencyResetRejected := GVL_HMI.uiIoEmergencyResult <> UINT#1;
    GVL_HMI.udiIoEmergencyAckSeq := udiIoEmergencyRequestSeq;
END_IF;
END_METHOD

METHOD PRIVATE ReadHmiCommands
// Request counters belong to gateway; pulses and acknowledgements belong to PLC.
udiHmiCommandNowMs := TIME_TO_UDINT(TIME());
GVL_HMI.udiHmiCommandClockMs := udiHmiCommandNowMs;
FOR uiHmiCommandIndex := UINT#1 TO UINT#121 DO
	axHmiCommandConsumed[uiHmiCommandIndex] := FALSE;
	axHmiCommandPulse[uiHmiCommandIndex] := FALSE;
	// Mandatory low scan rearms every existing R_TRIG, including scenario events.
	IF NOT axHmiCommandWasHigh[uiHmiCommandIndex] THEN
		IF axHmiInternalPulse[uiHmiCommandIndex] THEN
			axHmiCommandPulse[uiHmiCommandIndex] := TRUE;
			axHmiInternalPulse[uiHmiCommandIndex] := FALSE;
		ELSE
			audiHmiCommandSnapshot[uiHmiCommandIndex] := GVL_HMI.audiHmiCommandSeq[uiHmiCommandIndex];
			IF (audiHmiCommandSnapshot[uiHmiCommandIndex] <> UDINT#0)
			AND (audiHmiCommandSnapshot[uiHmiCommandIndex] <> GVL_HMI.audiHmiCommandAckSeq[uiHmiCommandIndex]) THEN
				axHmiCommandConsumed[uiHmiCommandIndex] := TRUE;
				IF IsHmiCommandFresh(udiIssuedAtMs := GVL_HMI.audiHmiCommandIssuedAtMs[uiHmiCommandIndex]) THEN
					axHmiCommandPulse[uiHmiCommandIndex] := TRUE;
					GVL_HMI.auiHmiCommandResult[uiHmiCommandIndex] := UINT#1;
				ELSE
					GVL_HMI.auiHmiCommandResult[uiHmiCommandIndex] := UINT#2;
				END_IF;
			END_IF;
		END_IF;
	END_IF;
	axHmiCommandWasHigh[uiHmiCommandIndex] := axHmiCommandPulse[uiHmiCommandIndex];
END_FOR;

// Stable wire IDs; command-contract.mjs and static tests enforce this mapping.
GVL_HMI.xCellEnable := axHmiCommandPulse[1];
GVL_HMI.xCellDisable := axHmiCommandPulse[2];
GVL_HMI.xCellStart := axHmiCommandPulse[3];
GVL_HMI.xCellStop := axHmiCommandPulse[4];
GVL_HMI.xCellReset := axHmiCommandPulse[5];
GVL_HMI.xSafetyRelayReset := axHmiCommandPulse[6];
GVL_HMI.xCellOperatorCancel := axHmiCommandPulse[7];
GVL_HMI.xAlarmResetWarnings := axHmiCommandPulse[8];
GVL_HMI.xModbusSettingsApply := axHmiCommandPulse[9];
GVL_HMI.stMultiType.Command.xAutoDistribute := axHmiCommandPulse[10];
GVL_HMI.xSimAxisGroupError := axHmiCommandPulse[11];
GVL_HMI.xSimRobotWrongAction := axHmiCommandPulse[12];
GVL_HMI.xSimCellBothGrippers := axHmiCommandPulse[13];
GVL_HMI.xSimPointXOutOfLimit := axHmiCommandPulse[14];
GVL_HMI.xSimPointYOutOfLimit := axHmiCommandPulse[15];
GVL_HMI.xSimPointZOutOfLimit := axHmiCommandPulse[16];
GVL_HMI.xSimPointInvalidVelocity := axHmiCommandPulse[17];
GVL_HMI.xSimMagazineWrongOperation := axHmiCommandPulse[18];
GVL_HMI.xSimMagazineNoBlank := axHmiCommandPulse[19];
GVL_HMI.xSimMagazineNoFreeSlot := axHmiCommandPulse[20];
GVL_HMI.xSimMagazineInvalidSlot := axHmiCommandPulse[21];
GVL_HMI.xSimMagazineSlotContent := axHmiCommandPulse[22];
GVL_HMI.xSimMagazineGeometry := axHmiCommandPulse[23];
GVL_HMI.xRobotDrivesEnable := axHmiCommandPulse[24];
GVL_HMI.xRobotDrivesDisable := axHmiCommandPulse[25];
GVL_HMI.xRobotStop := axHmiCommandPulse[26];
GVL_HMI.xRobotReset := axHmiCommandPulse[27];
GVL_HMI.xTestEnvironmentApply := axHmiCommandPulse[28];
GVL_HMI.xTestSpeedProfileApply := axHmiCommandPulse[29];
GVL_HMI.xTestScenarioApply := axHmiCommandPulse[30];
GVL_HMI.xPointCheckStop := axHmiCommandPulse[31];
GVL_HMI.xRobotManualExecute := axHmiCommandPulse[32];
GVL_HMI.stMultiType.Command.xSetTypeCount := axHmiCommandPulse[33];
GVL_HMI.xCellOperatorChoice := axHmiCommandPulse[34];
GVL_HMI.stMultiType.Command.xSetMachineType := axHmiCommandPulse[35];
GVL_HMI.xRobotControlModeApply := axHmiCommandPulse[36];
GVL_HMI.stMultiType.Command.xSetSlotType := axHmiCommandPulse[37];
GVL_HMI.astAxisHmiCommand[1].xHome := axHmiCommandPulse[38];
GVL_HMI.astAxisHmiCommand[1].xMoveAbsolute := axHmiCommandPulse[39];
GVL_HMI.astAxisHmiCommand[1].xMoveRelative := axHmiCommandPulse[40];
GVL_HMI.axSimAxisJogConflict[1] := axHmiCommandPulse[41];
GVL_HMI.axMachineSimReset[1] := axHmiCommandPulse[42];
GVL_HMI.axMachineEnable[1] := axHmiCommandPulse[43];
GVL_HMI.axMachineDisable[1] := axHmiCommandPulse[44];
GVL_HMI.axMachineReset[1] := axHmiCommandPulse[45];
GVL_HMI.axMachineSetBlank[1] := axHmiCommandPulse[46];
GVL_HMI.axMachineSetDetail[1] := axHmiCommandPulse[47];
GVL_HMI.axMachineAcceptDoor[1] := axHmiCommandPulse[48];
GVL_HMI.axMachineRejectDoor[1] := axHmiCommandPulse[49];
GVL_HMI.axMachineAcceptRun[1] := axHmiCommandPulse[50];
GVL_HMI.axMachineRejectRun[1] := axHmiCommandPulse[51];
GVL_HMI.axMachineManualSafetyDoorOpen[1] := axHmiCommandPulse[52];
GVL_HMI.axMachineManualSafetyDoorClose[1] := axHmiCommandPulse[53];
GVL_HMI.axMachineManualHatchOpen[1] := axHmiCommandPulse[54];
GVL_HMI.axMachineManualHatchClose[1] := axHmiCommandPulse[55];
GVL_HMI.axMachineManualHatchUnlock[1] := axHmiCommandPulse[56];
GVL_HMI.axMachineManualHatchLock[1] := axHmiCommandPulse[57];
GVL_HMI.axMachineManualChuckOpen[1] := axHmiCommandPulse[58];
GVL_HMI.axMachineManualChuckClose[1] := axHmiCommandPulse[59];
GVL_HMI.astAxisHmiCommand[2].xHome := axHmiCommandPulse[60];
GVL_HMI.astAxisHmiCommand[2].xMoveAbsolute := axHmiCommandPulse[61];
GVL_HMI.astAxisHmiCommand[2].xMoveRelative := axHmiCommandPulse[62];
GVL_HMI.axSimAxisJogConflict[2] := axHmiCommandPulse[63];
GVL_HMI.axMachineSimReset[2] := axHmiCommandPulse[64];
GVL_HMI.axMachineEnable[2] := axHmiCommandPulse[65];
GVL_HMI.axMachineDisable[2] := axHmiCommandPulse[66];
GVL_HMI.axMachineReset[2] := axHmiCommandPulse[67];
GVL_HMI.axMachineSetBlank[2] := axHmiCommandPulse[68];
GVL_HMI.axMachineSetDetail[2] := axHmiCommandPulse[69];
GVL_HMI.axMachineAcceptDoor[2] := axHmiCommandPulse[70];
GVL_HMI.axMachineRejectDoor[2] := axHmiCommandPulse[71];
GVL_HMI.axMachineAcceptRun[2] := axHmiCommandPulse[72];
GVL_HMI.axMachineRejectRun[2] := axHmiCommandPulse[73];
GVL_HMI.axMachineManualSafetyDoorOpen[2] := axHmiCommandPulse[74];
GVL_HMI.axMachineManualSafetyDoorClose[2] := axHmiCommandPulse[75];
GVL_HMI.axMachineManualHatchOpen[2] := axHmiCommandPulse[76];
GVL_HMI.axMachineManualHatchClose[2] := axHmiCommandPulse[77];
GVL_HMI.axMachineManualHatchUnlock[2] := axHmiCommandPulse[78];
GVL_HMI.axMachineManualHatchLock[2] := axHmiCommandPulse[79];
GVL_HMI.axMachineManualChuckOpen[2] := axHmiCommandPulse[80];
GVL_HMI.axMachineManualChuckClose[2] := axHmiCommandPulse[81];
GVL_HMI.astAxisHmiCommand[3].xHome := axHmiCommandPulse[82];
GVL_HMI.astAxisHmiCommand[3].xMoveAbsolute := axHmiCommandPulse[83];
GVL_HMI.astAxisHmiCommand[3].xMoveRelative := axHmiCommandPulse[84];
GVL_HMI.axSimAxisJogConflict[3] := axHmiCommandPulse[85];
GVL_HMI.axMachineSimReset[3] := axHmiCommandPulse[86];
GVL_HMI.axMachineEnable[3] := axHmiCommandPulse[87];
GVL_HMI.axMachineDisable[3] := axHmiCommandPulse[88];
GVL_HMI.axMachineReset[3] := axHmiCommandPulse[89];
GVL_HMI.axMachineSetBlank[3] := axHmiCommandPulse[90];
GVL_HMI.axMachineSetDetail[3] := axHmiCommandPulse[91];
GVL_HMI.axMachineAcceptDoor[3] := axHmiCommandPulse[92];
GVL_HMI.axMachineRejectDoor[3] := axHmiCommandPulse[93];
GVL_HMI.axMachineAcceptRun[3] := axHmiCommandPulse[94];
GVL_HMI.axMachineRejectRun[3] := axHmiCommandPulse[95];
GVL_HMI.axMachineManualSafetyDoorOpen[3] := axHmiCommandPulse[96];
GVL_HMI.axMachineManualSafetyDoorClose[3] := axHmiCommandPulse[97];
GVL_HMI.axMachineManualHatchOpen[3] := axHmiCommandPulse[98];
GVL_HMI.axMachineManualHatchClose[3] := axHmiCommandPulse[99];
GVL_HMI.axMachineManualHatchUnlock[3] := axHmiCommandPulse[100];
GVL_HMI.axMachineManualHatchLock[3] := axHmiCommandPulse[101];
GVL_HMI.axMachineManualChuckOpen[3] := axHmiCommandPulse[102];
GVL_HMI.axMachineManualChuckClose[3] := axHmiCommandPulse[103];
GVL_HMI.astMagazineCommand[1].xEnable := axHmiCommandPulse[104];
GVL_HMI.astMagazineCommand[1].xDisable := axHmiCommandPulse[105];
GVL_HMI.astMagazineCommand[1].xStop := axHmiCommandPulse[106];
GVL_HMI.astMagazineCommand[1].xReset := axHmiCommandPulse[107];
GVL_HMI.astMagazineCommand[1].xFill := axHmiCommandPulse[108];
GVL_HMI.astMagazineCommand[1].xClear := axHmiCommandPulse[109];
GVL_HMI.astMagazineCommand[1].xApplySlot := axHmiCommandPulse[110];
GVL_HMI.astMagazineCommand[1].xApplyPitchX := axHmiCommandPulse[111];
GVL_HMI.astMagazineCommand[1].xApplyPitchY := axHmiCommandPulse[112];
GVL_HMI.astMagazineCommand[2].xEnable := axHmiCommandPulse[113];
GVL_HMI.astMagazineCommand[2].xDisable := axHmiCommandPulse[114];
GVL_HMI.astMagazineCommand[2].xStop := axHmiCommandPulse[115];
GVL_HMI.astMagazineCommand[2].xReset := axHmiCommandPulse[116];
GVL_HMI.astMagazineCommand[2].xFill := axHmiCommandPulse[117];
GVL_HMI.astMagazineCommand[2].xClear := axHmiCommandPulse[118];
GVL_HMI.astMagazineCommand[2].xApplySlot := axHmiCommandPulse[119];
GVL_HMI.astMagazineCommand[2].xApplyPitchX := axHmiCommandPulse[120];
GVL_HMI.astMagazineCommand[2].xApplyPitchY := axHmiCommandPulse[121];
END_METHOD

METHOD PRIVATE RunRobotModbus
// Эффективная конфигурация всегда принадлежит RETAIN-GVL. HMI меняет только
// подготовленные значения и затем выдаёт отдельный импульс Apply.
// Новые RETAIN-поля после Online Change могут прийти нулевыми — нормализуем их
// до безопасных штатных значений до первого использования FB_ROBOT.
IF (GVL_ROBOT_MODBUS_RETAIN.tCommandStartTimeout < T#1S)
OR (GVL_ROBOT_MODBUS_RETAIN.tCommandStartTimeout > T#600S) THEN
	GVL_ROBOT_MODBUS_RETAIN.tCommandStartTimeout := T#30S;
END_IF;
IF (GVL_ROBOT_MODBUS_RETAIN.tCommandTimeout < T#1S)
OR (GVL_ROBOT_MODBUS_RETAIN.tCommandTimeout > T#3600S) THEN
	GVL_ROBOT_MODBUS_RETAIN.tCommandTimeout := T#600S;
END_IF;
GVL_ROBOT_MODBUS.Config.aIpAddress := GVL_ROBOT_MODBUS_RETAIN.aIpAddress;
GVL_ROBOT_MODBUS.Config.uiPort := GVL_ROBOT_MODBUS_RETAIN.uiPort;
GVL_ROBOT_MODBUS.Config.uiUnitId := GVL_ROBOT_MODBUS_RETAIN.uiUnitId;
GVL_ROBOT_MODBUS.Config.tResponseTimeout := GVL_ROBOT_MODBUS_RETAIN.tResponseTimeout;
GVL_ROBOT_MODBUS.Config.tPollInterval := GVL_ROBOT_MODBUS_RETAIN.tPollInterval;
GVL_ROBOT_MODBUS.Config.tHeartbeatTimeout := GVL_ROBOT_MODBUS_RETAIN.tHeartbeatTimeout;
GVL_ROBOT_MODBUS.Config.tCommandTimeout := GVL_ROBOT_MODBUS_RETAIN.tCommandTimeout;
GVL_ROBOT_MODBUS.xModeActive :=
	GVL_ROBOT_MODBUS_RETAIN.eControlMode = E_ROBOT_CONTROL_MODE.MODBUS_TCP;
GVL_HMI.xModbusMode := GVL_ROBOT_MODBUS.xModeActive;

IF NOT xModbusHmiInitialized THEN
	GVL_HMI.uiRobotControlModeRequest := TO_UINT(GVL_ROBOT_MODBUS_RETAIN.eControlMode);
	GVL_HMI.uiModbusIpOctet1 := BYTE_TO_UINT(GVL_ROBOT_MODBUS_RETAIN.aIpAddress[0]);
	GVL_HMI.uiModbusIpOctet2 := BYTE_TO_UINT(GVL_ROBOT_MODBUS_RETAIN.aIpAddress[1]);
	GVL_HMI.uiModbusIpOctet3 := BYTE_TO_UINT(GVL_ROBOT_MODBUS_RETAIN.aIpAddress[2]);
	GVL_HMI.uiModbusIpOctet4 := BYTE_TO_UINT(GVL_ROBOT_MODBUS_RETAIN.aIpAddress[3]);
	GVL_HMI.uiModbusPort := GVL_ROBOT_MODBUS_RETAIN.uiPort;
	GVL_HMI.uiModbusUnitId := GVL_ROBOT_MODBUS_RETAIN.uiUnitId;
	GVL_HMI.udiModbusResponseTimeoutMs := TIME_TO_UDINT(GVL_ROBOT_MODBUS_RETAIN.tResponseTimeout);
	GVL_HMI.udiModbusPollIntervalMs := TIME_TO_UDINT(GVL_ROBOT_MODBUS_RETAIN.tPollInterval);
	GVL_HMI.udiModbusHeartbeatTimeoutMs := TIME_TO_UDINT(GVL_ROBOT_MODBUS_RETAIN.tHeartbeatTimeout);
	GVL_HMI.udiModbusCommandStartTimeoutMs := TIME_TO_UDINT(GVL_ROBOT_MODBUS_RETAIN.tCommandStartTimeout);
	GVL_HMI.udiModbusCommandTimeoutMs := TIME_TO_UDINT(GVL_ROBOT_MODBUS_RETAIN.tCommandTimeout);
	xModbusHmiInitialized := TRUE;
END_IF;

xAllMachinesIdle := NOT GVL_MACHINE.Status[1].xBusy
	AND NOT GVL_MACHINE.Status[2].xBusy
	AND NOT GVL_MACHINE.Status[3].xBusy;
xModeCommonSafe := xHmiConnectionAlive
	AND NOT GVL_CELL_MANAGER.Status.xRunning
	AND NOT GVL_MAGAZINE.astStatus[1].xBusy
	AND NOT GVL_MAGAZINE.astStatus[2].xBusy
	AND xAllMachinesIdle
	AND NOT GVL_ROBOT.Status.xBusy
	AND NOT GVL_HMI.xRobotManualExecute;

IF GVL_ROBOT_MODBUS.xModeActive THEN
	GVL_ROBOT_MODBUS.xRobotModeChangeAllowed := xModeCommonSafe
		AND GVL_ROBOT_MODBUS.Status.xCommunicationAlive
		AND (GVL_ROBOT_MODBUS.Status.uiExecutionState =
			TO_UINT(E_ROBOT_MODBUS_EXECUTION_STATE.IDLE))
		AND NOT GVL_ROBOT_MODBUS.Status.xDrivesEnabled;
ELSE
	GVL_ROBOT_MODBUS.xRobotModeChangeAllowed := xModeCommonSafe
		AND xDrivesOff
		AND NOT xMotionBusy
		AND GVL_ROBOT_MODBUS.Status.xConfigValid;
END_IF;

GVL_ROBOT_MODBUS.xSettingsChangeAllowed := xHmiConnectionAlive
	AND NOT GVL_CELL_MANAGER.Status.xRunning
	AND NOT GVL_MAGAZINE.astStatus[1].xBusy
	AND NOT GVL_MAGAZINE.astStatus[2].xBusy
	AND xAllMachinesIdle
	AND NOT GVL_ROBOT.Status.xBusy;

rtRobotModeApply(CLK := GVL_HMI.xRobotControlModeApply);
rtModbusSettingsApply(CLK := GVL_HMI.xModbusSettingsApply);
GVL_ROBOT_MODBUS.xReconnectRequest := FALSE;

IF rtModbusSettingsApply.Q THEN
	IF GVL_ROBOT_MODBUS.xSettingsChangeAllowed
	AND (GVL_HMI.uiModbusIpOctet1 >= UINT#1)
	AND (GVL_HMI.uiModbusIpOctet1 <= UINT#223)
	AND (GVL_HMI.uiModbusIpOctet2 <= UINT#255)
	AND (GVL_HMI.uiModbusIpOctet3 <= UINT#255)
	AND (GVL_HMI.uiModbusIpOctet4 <= UINT#255)
	AND (GVL_HMI.uiModbusPort >= UINT#1)
	AND (GVL_HMI.uiModbusUnitId <= UINT#255)
	AND (GVL_HMI.udiModbusResponseTimeoutMs >= UDINT#50)
	AND (GVL_HMI.udiModbusResponseTimeoutMs <= UDINT#10000)
	AND (GVL_HMI.udiModbusPollIntervalMs >= UDINT#10)
	AND (GVL_HMI.udiModbusPollIntervalMs <= UDINT#5000)
	AND (GVL_HMI.udiModbusHeartbeatTimeoutMs >= UDINT#500)
	AND (GVL_HMI.udiModbusHeartbeatTimeoutMs <= UDINT#30000)
	AND (GVL_HMI.udiModbusCommandStartTimeoutMs >= UDINT#1000)
	AND (GVL_HMI.udiModbusCommandStartTimeoutMs <= UDINT#600000)
	AND (GVL_HMI.udiModbusCommandTimeoutMs >= UDINT#1000)
	AND (GVL_HMI.udiModbusCommandTimeoutMs <= UDINT#3600000) THEN
		GVL_ROBOT_MODBUS_RETAIN.aIpAddress[0] := UINT_TO_BYTE(GVL_HMI.uiModbusIpOctet1);
		GVL_ROBOT_MODBUS_RETAIN.aIpAddress[1] := UINT_TO_BYTE(GVL_HMI.uiModbusIpOctet2);
		GVL_ROBOT_MODBUS_RETAIN.aIpAddress[2] := UINT_TO_BYTE(GVL_HMI.uiModbusIpOctet3);
		GVL_ROBOT_MODBUS_RETAIN.aIpAddress[3] := UINT_TO_BYTE(GVL_HMI.uiModbusIpOctet4);
		GVL_ROBOT_MODBUS_RETAIN.uiPort := GVL_HMI.uiModbusPort;
		GVL_ROBOT_MODBUS_RETAIN.uiUnitId := GVL_HMI.uiModbusUnitId;
		GVL_ROBOT_MODBUS_RETAIN.tResponseTimeout := UDINT_TO_TIME(GVL_HMI.udiModbusResponseTimeoutMs);
		GVL_ROBOT_MODBUS_RETAIN.tPollInterval := UDINT_TO_TIME(GVL_HMI.udiModbusPollIntervalMs);
		GVL_ROBOT_MODBUS_RETAIN.tHeartbeatTimeout := UDINT_TO_TIME(GVL_HMI.udiModbusHeartbeatTimeoutMs);
		GVL_ROBOT_MODBUS_RETAIN.tCommandStartTimeout := UDINT_TO_TIME(GVL_HMI.udiModbusCommandStartTimeoutMs);
		GVL_ROBOT_MODBUS_RETAIN.tCommandTimeout := UDINT_TO_TIME(GVL_HMI.udiModbusCommandTimeoutMs);
		GVL_ROBOT_MODBUS.xReconnectRequest := GVL_ROBOT_MODBUS.xModeActive;
		GVL_HMI.uiModbusSettingsRejectReason := UINT#0;
	ELSE
		GVL_HMI.uiModbusSettingsRejectReason := UINT#1;
		uiRobotInterfaceWarningCode := WRN_MODBUS_SETTINGS_REJECTED;
	END_IF;
END_IF;

IF rtRobotModeApply.Q THEN
	IF (GVL_HMI.uiRobotControlModeRequest <= UINT#1)
	AND GVL_ROBOT_MODBUS.xRobotModeChangeAllowed THEN
	IF GVL_HMI.uiRobotControlModeRequest = UINT#1 THEN
			GVL_ROBOT_MODBUS_RETAIN.eControlMode := E_ROBOT_CONTROL_MODE.MODBUS_TCP;
		ELSE
			GVL_ROBOT_MODBUS_RETAIN.eControlMode := E_ROBOT_CONTROL_MODE.SOFTMOTION;
		END_IF;
		GVL_HMI.uiRobotControlModeRequest := TO_UINT(GVL_ROBOT_MODBUS_RETAIN.eControlMode);
		GVL_HMI.uiRobotModeRejectReason := UINT#0;
	ELSE
		IF NOT xModeCommonSafe THEN
			GVL_HMI.uiRobotModeRejectReason := UINT#1;
		ELSIF NOT GVL_ROBOT_MODBUS.xModeActive AND NOT xDrivesOff THEN
			GVL_HMI.uiRobotModeRejectReason := UINT#2;
		ELSIF GVL_ROBOT_MODBUS.xModeActive THEN
			GVL_HMI.uiRobotModeRejectReason := UINT#3;
		ELSE
			GVL_HMI.uiRobotModeRejectReason := UINT#4;
		END_IF;
		uiRobotInterfaceWarningCode := WRN_ROBOT_MODE_REJECTED;
		GVL_HMI.uiRobotControlModeRequest := TO_UINT(GVL_ROBOT_MODBUS_RETAIN.eControlMode);
	END_IF;
END_IF;

// Повторная выборка после возможного Apply исключает один цикл старого режима.
GVL_ROBOT_MODBUS.xModeActive :=
	GVL_ROBOT_MODBUS_RETAIN.eControlMode = E_ROBOT_CONTROL_MODE.MODBUS_TCP;
GVL_HMI.xModbusMode := GVL_ROBOT_MODBUS.xModeActive;
GVL_ROBOT_MODBUS.Config.aIpAddress := GVL_ROBOT_MODBUS_RETAIN.aIpAddress;
GVL_ROBOT_MODBUS.Config.uiPort := GVL_ROBOT_MODBUS_RETAIN.uiPort;
GVL_ROBOT_MODBUS.Config.uiUnitId := GVL_ROBOT_MODBUS_RETAIN.uiUnitId;
GVL_ROBOT_MODBUS.Config.tResponseTimeout := GVL_ROBOT_MODBUS_RETAIN.tResponseTimeout;
GVL_ROBOT_MODBUS.Config.tPollInterval := GVL_ROBOT_MODBUS_RETAIN.tPollInterval;
GVL_ROBOT_MODBUS.Config.tHeartbeatTimeout := GVL_ROBOT_MODBUS_RETAIN.tHeartbeatTimeout;
GVL_ROBOT_MODBUS.Config.tCommandTimeout := GVL_ROBOT_MODBUS_RETAIN.tCommandTimeout;

ROBOT_MODBUS(
	xEnable := GVL_ROBOT_MODBUS.xModeActive,
	xReconnect := GVL_ROBOT_MODBUS.xReconnectRequest,
	Config := GVL_ROBOT_MODBUS.Config,
	Command := GVL_ROBOT.ModbusCommand,
	Status => GVL_ROBOT_MODBUS.Status,
	auiWriteRegisters := GVL_ROBOT_MODBUS.auiWriteRegisters,
	auiReadRegisters := GVL_ROBOT_MODBUS.auiReadRegisters
);

GVL_ROBOT.xModbusBusy := GVL_ROBOT_MODBUS.Status.xBusy;
GVL_ROBOT.xModbusDone := GVL_ROBOT_MODBUS.Status.xDone;
GVL_ROBOT.xModbusError := GVL_ROBOT_MODBUS.Status.xError;

IF GVL_ROBOT_MODBUS.xModeActive THEN
	xRobotInterfaceReady := GVL_ROBOT_MODBUS.Status.xReady;
	xDrivesReady := GVL_ROBOT_MODBUS.Status.xReady;
	xDrivesPowered := GVL_ROBOT_MODBUS.Status.xDrivesEnabled;
	xDrivesOff := NOT GVL_ROBOT_MODBUS.Status.xDrivesEnabled;
	xPowerTransitionActive := FALSE;
	xMotionBusy := GVL_ROBOT_MODBUS.Status.xBusy;
	xDriveError := GVL_ROBOT_MODBUS.Status.xError;
	lrRobotActualX := GVL_ROBOT_MODBUS.Status.lrActualX;
	lrRobotActualY := GVL_ROBOT_MODBUS.Status.lrActualY;
	lrRobotActualZ := GVL_ROBOT_MODBUS.Status.lrActualZ;
	GVL_HMI.lrActualX := lrRobotActualX;
	GVL_HMI.lrActualY := lrRobotActualY;
	GVL_HMI.lrActualZ := lrRobotActualZ;
	GVL_HMI.HMI.ActualX := lrRobotActualX;
	GVL_HMI.HMI.ActualY := lrRobotActualY;
	GVL_HMI.HMI.ActualZ := lrRobotActualZ;
ELSE
	xRobotInterfaceReady := TRUE;
	// Не публикуем просроченные Modbus-координаты: в SoftMotion активен только
	// локальный источник обратной связи.
	GVL_ROBOT_MODBUS.Status.lrActualX := LREAL#0.0;
	GVL_ROBOT_MODBUS.Status.lrActualY := LREAL#0.0;
	GVL_ROBOT_MODBUS.Status.lrActualZ := LREAL#0.0;
	lrRobotActualX := GVL_AXIS_GROUP.AxisGroup.Status.ActualX;
	lrRobotActualY := GVL_AXIS_GROUP.AxisGroup.Status.ActualY;
	lrRobotActualZ := GVL_AXIS_GROUP.AxisGroup.Status.ActualZ;
END_IF;
END_METHOD

METHOD PRIVATE RunRobot
// Старый типизированный канал сохраняется для совместимости. Новый HMI пишет
// числовые коды, которые преобразуются в enum только внутри PLC.
stRobotHmiCommand := GVL_HMI.stRobotCommand;
xHmiRobotActionAttempt := GVL_HMI.xRobotManualExecute OR GVL_HMI.stRobotCommand.xExecute;

// Числовой канал HMI хранит последнюю отправленную команду, а не текущий выбор
// в интерфейсе. Разрешение её цели используется только в скане попытки запуска;
// между запросами HMI получает общее разрешение ручного движения.
// Типизированный legacy-канал остаётся владельцем своей команды при прямом Execute.
eHmiRobotStatusAction := stRobotHmiCommand.eAction;
eHmiRobotStatusPoint := stRobotHmiCommand.eSetPoint;
IF GVL_HMI.uiRobotManualAction > UINT#0 THEN
	CASE GVL_HMI.uiRobotManualAction OF
		1: eHmiRobotStatusAction := E_ROBOT_ACTION.MOVE_TO_POINT;
		2: eHmiRobotStatusAction := E_ROBOT_ACTION.UNCLAMP_1;
		3: eHmiRobotStatusAction := E_ROBOT_ACTION.CLAMP_1;
		4: eHmiRobotStatusAction := E_ROBOT_ACTION.UNCLAMP_2;
		5: eHmiRobotStatusAction := E_ROBOT_ACTION.CLAMP_2;
		6: eHmiRobotStatusAction := E_ROBOT_ACTION.ROTATE_TO_BLANK;
		7: eHmiRobotStatusAction := E_ROBOT_ACTION.ROTATE_TO_DETAIL;
	ELSE
		eHmiRobotStatusAction := E_ROBOT_ACTION.NONE;
	END_CASE;
	CASE GVL_HMI.uiRobotManualPoint OF
		1: eHmiRobotStatusPoint := E_POINT_NAME.MACHINE_1_ABOVE;
		3: eHmiRobotStatusPoint := E_POINT_NAME.MACHINE_1_CHUCK_APROACH;
		4: eHmiRobotStatusPoint := E_POINT_NAME.MACHINE_1_CHUCK_POSITION;
		5: eHmiRobotStatusPoint := E_POINT_NAME.MACHINE_2_ABOVE;
		7: eHmiRobotStatusPoint := E_POINT_NAME.MACHINE_2_CHUCK_APROACH;
		8: eHmiRobotStatusPoint := E_POINT_NAME.MACHINE_2_CHUCK_POSITION;
		9: eHmiRobotStatusPoint := E_POINT_NAME.MACHINE_3_ABOVE;
		11: eHmiRobotStatusPoint := E_POINT_NAME.MACHINE_3_CHUCK_APROACH;
		12: eHmiRobotStatusPoint := E_POINT_NAME.MACHINE_3_CHUCK_POSITION;
		13: eHmiRobotStatusPoint := E_POINT_NAME.HOME_SAFETY;
		14: eHmiRobotStatusPoint := E_POINT_NAME.MAGAZINE_SAFE;
		15: eHmiRobotStatusPoint := E_POINT_NAME.MAGAZINE_CHANGE;
		16: eHmiRobotStatusPoint := E_POINT_NAME.MAGAZINE_IN_SLOT;
		17: eHmiRobotStatusPoint := E_POINT_NAME.GEOMETRY_1_SAFE;
		18: eHmiRobotStatusPoint := E_POINT_NAME.GEOMETRY_1_CHANGE;
		19: eHmiRobotStatusPoint := E_POINT_NAME.GEOMETRY_1_PLACE;
		20: eHmiRobotStatusPoint := E_POINT_NAME.GEOMETRY_2_SAFE;
		21: eHmiRobotStatusPoint := E_POINT_NAME.GEOMETRY_2_CHANGE;
		22: eHmiRobotStatusPoint := E_POINT_NAME.GEOMETRY_2_PLACE;
	ELSE
		eHmiRobotStatusPoint := E_POINT_NAME.NONE;
	END_CASE;
END_IF;

IF GVL_HMI.xRobotManualExecute THEN
	stRobotHmiCommand.xExecute := FALSE;
	stRobotHmiCommand.eAction := E_ROBOT_ACTION.NONE;
	stRobotHmiCommand.eSetPoint := E_POINT_NAME.NONE;
	CASE GVL_HMI.uiRobotManualAction OF
		1: stRobotHmiCommand.eAction := E_ROBOT_ACTION.MOVE_TO_POINT;
		2: stRobotHmiCommand.eAction := E_ROBOT_ACTION.UNCLAMP_1;
		3: stRobotHmiCommand.eAction := E_ROBOT_ACTION.CLAMP_1;
		4: stRobotHmiCommand.eAction := E_ROBOT_ACTION.UNCLAMP_2;
		5: stRobotHmiCommand.eAction := E_ROBOT_ACTION.CLAMP_2;
		6: stRobotHmiCommand.eAction := E_ROBOT_ACTION.ROTATE_TO_BLANK;
		7: stRobotHmiCommand.eAction := E_ROBOT_ACTION.ROTATE_TO_DETAIL;
	END_CASE;
	CASE GVL_HMI.uiRobotManualPoint OF
		1: stRobotHmiCommand.eSetPoint := E_POINT_NAME.MACHINE_1_ABOVE;
		3: stRobotHmiCommand.eSetPoint := E_POINT_NAME.MACHINE_1_CHUCK_APROACH;
		4: stRobotHmiCommand.eSetPoint := E_POINT_NAME.MACHINE_1_CHUCK_POSITION;
		5: stRobotHmiCommand.eSetPoint := E_POINT_NAME.MACHINE_2_ABOVE;
		7: stRobotHmiCommand.eSetPoint := E_POINT_NAME.MACHINE_2_CHUCK_APROACH;
		8: stRobotHmiCommand.eSetPoint := E_POINT_NAME.MACHINE_2_CHUCK_POSITION;
		9: stRobotHmiCommand.eSetPoint := E_POINT_NAME.MACHINE_3_ABOVE;
		11: stRobotHmiCommand.eSetPoint := E_POINT_NAME.MACHINE_3_CHUCK_APROACH;
		12: stRobotHmiCommand.eSetPoint := E_POINT_NAME.MACHINE_3_CHUCK_POSITION;
		13: stRobotHmiCommand.eSetPoint := E_POINT_NAME.HOME_SAFETY;
		14: stRobotHmiCommand.eSetPoint := E_POINT_NAME.MAGAZINE_SAFE;
		15: stRobotHmiCommand.eSetPoint := E_POINT_NAME.MAGAZINE_CHANGE;
		16: stRobotHmiCommand.eSetPoint := E_POINT_NAME.MAGAZINE_IN_SLOT;
		17: stRobotHmiCommand.eSetPoint := E_POINT_NAME.GEOMETRY_1_SAFE;
		18: stRobotHmiCommand.eSetPoint := E_POINT_NAME.GEOMETRY_1_CHANGE;
		19: stRobotHmiCommand.eSetPoint := E_POINT_NAME.GEOMETRY_1_PLACE;
		20: stRobotHmiCommand.eSetPoint := E_POINT_NAME.GEOMETRY_2_SAFE;
		21: stRobotHmiCommand.eSetPoint := E_POINT_NAME.GEOMETRY_2_CHANGE;
		22: stRobotHmiCommand.eSetPoint := E_POINT_NAME.GEOMETRY_2_PLACE;
	END_CASE;
	IF GVL_HMI.uiRobotManualSlot <= SINT_TO_UINT(GVL_CELL_SETTINGS.NumberDetail) THEN
		stRobotHmiCommand.iActiveSlot := UINT_TO_SINT(GVL_HMI.uiRobotManualSlot);
	ELSE
		stRobotHmiCommand.iActiveSlot := SINT#0;
	END_IF;
	stRobotHmiCommand.uiMagazineId := GVL_HMI.uiRobotManualMagazine;
END_IF;

// Два FB_MAGAZINE не имеют права одновременно владеть роботом.
stSelectedMagazineCommand.xExecute := FALSE;
stSelectedMagazineCommand.xStop := FALSE;
stSelectedMagazineCommand.xReset := FALSE;
stSelectedMagazineCommand.eAction := E_ROBOT_ACTION.NONE;
stSelectedMagazineCommand.eSetPoint := E_POINT_NAME.NONE;
stSelectedMagazineCommand.iActiveSlot := SINT#0;
stSelectedMagazineCommand.uiMagazineId := UINT#0;
IF GVL_MAGAZINE.astCommand[1].xExecute OR GVL_MAGAZINE.astCommand[1].xStop THEN
	stSelectedMagazineCommand := GVL_MAGAZINE.astCommand[1];
ELSIF GVL_MAGAZINE.astCommand[2].xExecute OR GVL_MAGAZINE.astCommand[2].xStop THEN
	stSelectedMagazineCommand := GVL_MAGAZINE.astCommand[2];
END_IF;

xHmiRobotActionBaseAllowed := xRobotHmiPermit
	AND NOT xPointCheckActive
	AND xHmiConnectionAlive
	AND NOT GVL_CELL_CONTROL.xGlobalError
	AND NOT GVL_ROBOT.Status.xBusy
	AND NOT GVL_ROBOT.Status.xError
	AND (GVL_ROBOT.Diag.eState = E_ROBOT_STATE.IDLE)
	AND (GVL_HMI.xModbusMode
		OR (GVL_MOTION_MANAGER.stMotionManager.Diag.eState = E_MOTION_MANAGER_STATE.IDLE))
	AND (
		(GVL_HMI.xModbusMode AND GVL_ROBOT_MODBUS.Status.xReady)
		OR (NOT GVL_HMI.xModbusMode
			AND xDrivesReady
			AND NOT xMotionBusy
			AND NOT xDriveError
			AND GVL_POINT_MANAGER.PointManager.Diag.xXLimitValid
			AND GVL_POINT_MANAGER.PointManager.Diag.xYLimitValid
			AND GVL_POINT_MANAGER.PointManager.Diag.xZLimitValid)
	);

// Ручное движение не зависит от готовности оборудования назначения.
// Единственное условие оборудования — подтверждённо открытый люк при входе
// внутрь станка. Оно одинаково для числового и legacy-канала.
xHmiRobotPointTargetAllowed := TRUE;
CASE stRobotHmiCommand.eSetPoint OF
	E_POINT_NAME.MACHINE_1_INSIDE,
	E_POINT_NAME.MACHINE_1_CHUCK_APROACH,
	E_POINT_NAME.MACHINE_1_CHUCK_POSITION:
		xHmiRobotPointTargetAllowed := GVL_MACHINE.Status[1].stIo.xDoorOpen
			AND NOT GVL_MACHINE.Status[1].stIo.xDoorClosed;
	E_POINT_NAME.MACHINE_2_INSIDE,
	E_POINT_NAME.MACHINE_2_CHUCK_APROACH,
	E_POINT_NAME.MACHINE_2_CHUCK_POSITION:
		xHmiRobotPointTargetAllowed := GVL_MACHINE.Status[2].stIo.xDoorOpen
			AND NOT GVL_MACHINE.Status[2].stIo.xDoorClosed;
	E_POINT_NAME.MACHINE_3_INSIDE,
	E_POINT_NAME.MACHINE_3_CHUCK_APROACH,
	E_POINT_NAME.MACHINE_3_CHUCK_POSITION:
		xHmiRobotPointTargetAllowed := GVL_MACHINE.Status[3].stIo.xDoorOpen
			AND NOT GVL_MACHINE.Status[3].stIo.xDoorClosed;
END_CASE;

xHmiRobotPointAllowed := xHmiRobotActionBaseAllowed
	AND (stRobotHmiCommand.eSetPoint <> E_POINT_NAME.NONE)
	AND xHmiRobotPointTargetAllowed
	AND (
		((stRobotHmiCommand.eSetPoint <> E_POINT_NAME.MAGAZINE_SAFE)
		AND (stRobotHmiCommand.eSetPoint <> E_POINT_NAME.MAGAZINE_CHANGE)
		AND (stRobotHmiCommand.eSetPoint <> E_POINT_NAME.MAGAZINE_IN_SLOT))
		OR (
			(stRobotHmiCommand.iActiveSlot >= SINT#1)
			AND (SINT_TO_UINT(stRobotHmiCommand.iActiveSlot)
				<= (GVL_CELL_SETTINGS.MagazineRows * GVL_CELL_SETTINGS.MagazineColumns))
			AND (stRobotHmiCommand.uiMagazineId >= UINT#1)
			AND (stRobotHmiCommand.uiMagazineId <= UINT#2)
		)
	);

// Захваты не зависят от питания и состояния Motion-слоя. В ручном режиме ими
// можно пользоваться при любой внешней аварии, пока исправен сам блок захвата
// и он не выполняет предыдущее действие.
xHmiGripperActionBaseAllowed := xRobotHmiPermit
	AND NOT xPointCheckActive
	AND xHmiConnectionAlive
	AND NOT GVL_ROBOT.Status.xBusy
	AND ((GVL_ROBOT.Diag.eState = E_ROBOT_STATE.IDLE)
		OR (NOT GVL_HMI.xModbusMode AND (GVL_ROBOT.Diag.eState = E_ROBOT_STATE.ERROR)))
	AND (
		(GVL_HMI.xModbusMode AND GVL_ROBOT_MODBUS.Status.xReady)
		OR (NOT GVL_HMI.xModbusMode
			AND (GVL_ROBOT.GripperError.dwAlarmActive = DWORD#0)
			AND (GVL_ROBOT.GripperDiag.eState = E_GRIPPER_STATE.IDLE))
	);

xHmiRobotActionAllowed := FALSE;
CASE stRobotHmiCommand.eAction OF
	E_ROBOT_ACTION.MOVE_TO_POINT:
		xHmiRobotActionAllowed := xHmiRobotPointAllowed;
	E_ROBOT_ACTION.UNCLAMP_1:
		xHmiRobotActionAllowed := xHmiGripperActionBaseAllowed
			AND NOT GVL_ROBOT.Status.xGripper1Open;
	E_ROBOT_ACTION.CLAMP_1:
		xHmiRobotActionAllowed := xHmiGripperActionBaseAllowed
			AND NOT GVL_ROBOT.Status.xGripper1Closed;
	E_ROBOT_ACTION.UNCLAMP_2:
		xHmiRobotActionAllowed := xHmiGripperActionBaseAllowed
			AND NOT GVL_ROBOT.Status.xGripper2Open;
	E_ROBOT_ACTION.CLAMP_2:
		xHmiRobotActionAllowed := xHmiGripperActionBaseAllowed
			AND NOT GVL_ROBOT.Status.xGripper2Closed;
	E_ROBOT_ACTION.ROTATE_TO_BLANK:
		xHmiRobotActionAllowed := xHmiGripperActionBaseAllowed
			AND NOT GVL_ROBOT.Status.xRotatedToBlank;
	E_ROBOT_ACTION.ROTATE_TO_DETAIL:
		xHmiRobotActionAllowed := xHmiGripperActionBaseAllowed
			AND NOT GVL_ROBOT.Status.xRotatedToDetail;
END_CASE;

IF GVL_HMI.xRobotManualExecute THEN
	stRobotHmiCommand.xExecute := xHmiRobotActionAllowed;
ELSIF stRobotHmiCommand.xExecute AND NOT xHmiRobotActionAllowed THEN
	stRobotHmiCommand.xExecute := FALSE;
END_IF;

// Общая ошибка запрещает координатное движение, но не ручное управление
// независимым пневматическим захватом.
IF GVL_CELL_CONTROL.xGlobalError
AND (stRobotHmiCommand.eAction = E_ROBOT_ACTION.MOVE_TO_POINT) THEN
	stRobotHmiCommand.xExecute := FALSE;
	stRobotHmiCommand.eAction := E_ROBOT_ACTION.NONE;
	stRobotHmiCommand.eSetPoint := E_POINT_NAME.NONE;
END_IF;
// Stop является импульсом текущего цикла и не должен защёлкиваться в локальной команде.
stRobotHmiCommand.xStop := xHmiStopAccepted;
rtHmiRobotAction(CLK := xHmiRobotActionAttempt);

// Единственный владелец временных точек разрешает координаты и для ручной,
// и для автоматической команды. FB_MAGAZINE больше не пишет общую таблицу.
stMagazinePointCommand := stSelectedMagazineCommand;
IF (stRobotHmiCommand.eSetPoint = E_POINT_NAME.MAGAZINE_SAFE)
OR (stRobotHmiCommand.eSetPoint = E_POINT_NAME.MAGAZINE_CHANGE)
OR (stRobotHmiCommand.eSetPoint = E_POINT_NAME.MAGAZINE_IN_SLOT) THEN
	stMagazinePointCommand := stRobotHmiCommand;
END_IF;
eMagazineBasePoint := E_POINT_NAME.NONE;
CASE stMagazinePointCommand.uiMagazineId OF
	UINT#1: eMagazineBasePoint := E_POINT_NAME.MAGAZINE_1_DETAIL;
	UINT#2: eMagazineBasePoint := E_POINT_NAME.MAGAZINE_2_DETAIL;
END_CASE;

IF NOT GVL_HMI.xModbusMode
AND (GVL_CELL_SETTINGS.MagazineRows > UINT#0)
AND (GVL_CELL_SETTINGS.MagazineColumns > UINT#0)
AND (eMagazineBasePoint <> E_POINT_NAME.NONE)
AND (stMagazinePointCommand.iActiveSlot >= SINT#1)
AND (SINT_TO_UINT(stMagazinePointCommand.iActiveSlot)
	<= (GVL_CELL_SETTINGS.MagazineRows * GVL_CELL_SETTINGS.MagazineColumns))
AND ((stMagazinePointCommand.eSetPoint = E_POINT_NAME.MAGAZINE_SAFE)
	OR (stMagazinePointCommand.eSetPoint = E_POINT_NAME.MAGAZINE_CHANGE)
	OR (stMagazinePointCommand.eSetPoint = E_POINT_NAME.MAGAZINE_IN_SLOT)) THEN
	uiRobotManualMagazineIndex := SINT_TO_UINT(stMagazinePointCommand.iActiveSlot - SINT#1);
	uiRobotManualMagazineColumn := uiRobotManualMagazineIndex MOD GVL_CELL_SETTINGS.MagazineColumns;
	uiRobotManualMagazineRow := uiRobotManualMagazineIndex / GVL_CELL_SETTINGS.MagazineColumns;
	GVL_POINT.Points[stMagazinePointCommand.eSetPoint] := GVL_POINT.Points[eMagazineBasePoint];
	GVL_POINT.Points[stMagazinePointCommand.eSetPoint].X :=
		GVL_POINT.Points[stMagazinePointCommand.eSetPoint].X
		+ UINT_TO_LREAL(uiRobotManualMagazineColumn) * GVL_HMI.MagazinePitchX;
	GVL_POINT.Points[stMagazinePointCommand.eSetPoint].Y :=
		GVL_POINT.Points[stMagazinePointCommand.eSetPoint].Y
		+ UINT_TO_LREAL(uiRobotManualMagazineRow) * GVL_HMI.MagazinePitchY;
	// Signed-смещение добавляется к базе: отрицательное Z поднимает траверсу, положительное опускает.
	IF stMagazinePointCommand.eSetPoint = E_POINT_NAME.MAGAZINE_SAFE THEN
		GVL_POINT.Points[stMagazinePointCommand.eSetPoint].Z :=
			GVL_POINT.Points[eMagazineBasePoint].Z
			+ GVL_POINT.Points[eMagazineBasePoint].MagazineSafeZ;
	ELSIF stMagazinePointCommand.eSetPoint = E_POINT_NAME.MAGAZINE_CHANGE THEN
		GVL_POINT.Points[stMagazinePointCommand.eSetPoint].Z :=
			GVL_POINT.Points[eMagazineBasePoint].Z
			+ GVL_POINT.Points[eMagazineBasePoint].MagazineChangeZ;
	END_IF;
END_IF;

// Внешний контроллер включается только со своего пульта. Из HMI доступны Stop,
// Reset и семантические команды при подтверждённой связи/готовности.
IF GVL_HMI.xModbusMode THEN
	GVL_HMI.stRobotHmiStatus.xDrivesPowered := GVL_ROBOT_MODBUS.Status.xDrivesEnabled;
	GVL_HMI.stRobotHmiStatus.xDrivesOff := NOT GVL_ROBOT_MODBUS.Status.xDrivesEnabled;
	GVL_HMI.stRobotHmiStatus.xPowerTransitionActive := FALSE;
	GVL_HMI.stRobotHmiStatus.xDrivesEnableAllowed := FALSE;
	GVL_HMI.stRobotHmiStatus.xDrivesDisableAllowed := FALSE;
	GVL_HMI.stRobotHmiStatus.xStopAllowed := xRobotHmiPermit
		AND GVL_ROBOT_MODBUS.Status.xCommunicationAlive
		AND GVL_ROBOT_MODBUS.Status.xBusy;
	GVL_HMI.stRobotHmiStatus.xResetAllowed := xRobotHmiPermit
		AND GVL_ROBOT_MODBUS.Status.xCommunicationAlive
		AND NOT GVL_ROBOT_MODBUS.Status.xBusy
		AND GVL_ROBOT_MODBUS.Status.xError;
	xHmiStopAccepted := GVL_HMI.xRobotStop
		AND GVL_HMI.stRobotHmiStatus.xStopAllowed;
END_IF;

// Отдельный владелец проверки инженерной точки. Все технологические условия
// вычисляются здесь, а мобильный клиент получает только результат xAllowed.
FOR uiPointCheckLoop := UINT#1 TO INT_TO_UINT(GVL_POINT.iEditablePointCount) DO
	stPointCheckCandidate := GVL_POINT.Points[aePointCheckNames[uiPointCheckLoop]];
	uiPointCheckReason := UINT#0;
	uiPointCheckMachine := UINT#0;
	IF (uiPointCheckLoop <= UINT#9) AND ((uiPointCheckLoop MOD UINT#3) <> UINT#1) THEN
		uiPointCheckMachine := (uiPointCheckLoop - UINT#1) / UINT#3 + UINT#1;
	END_IF;
	IF NOT xHmiConnectionAlive THEN
		uiPointCheckReason := UINT#3;
	ELSIF NOT GVL_CELL_CONTROL.xManual THEN
		uiPointCheckReason := UINT#4;
	ELSIF GVL_HMI.xModbusMode THEN
		uiPointCheckReason := UINT#5;
	ELSIF GVL_CELL_MANAGER.Status.xRunning THEN
		uiPointCheckReason := UINT#6;
	ELSIF GVL_CELL_CONTROL.xGlobalError THEN
		uiPointCheckReason := UINT#7;
	ELSIF xPointCheckActive OR GVL_ROBOT.Status.xBusy
	OR ((GVL_ROBOT.Diag.eState <> E_ROBOT_STATE.IDLE)
		AND (GVL_ROBOT.Diag.eState <> E_ROBOT_STATE.ERROR)) THEN
		uiPointCheckReason := UINT#8;
	ELSIF xMotionBusy
	OR ((GVL_MOTION_MANAGER.stMotionManager.Diag.eState <> E_MOTION_MANAGER_STATE.IDLE)
		AND (GVL_MOTION_MANAGER.stMotionManager.Diag.eState <> E_MOTION_MANAGER_STATE.ERROR)) THEN
		uiPointCheckReason := UINT#9;
	ELSIF xDriveError OR GVL_ROBOT.Status.xError OR GVL_MOTION_MANAGER.stMotionManager.Status.xError THEN
		uiPointCheckReason := UINT#10;
	ELSIF NOT xPointEditorAllHomed THEN
		uiPointCheckReason := UINT#11;
	ELSIF NOT GVL_AXIS_GROUP.AxisGroup.Status.xPositionValid THEN
		uiPointCheckReason := UINT#12;
	ELSIF NOT GVL_POINT_MANAGER.PointManager.Diag.xXLimitValid
	OR NOT GVL_POINT_MANAGER.PointManager.Diag.xYLimitValid
	OR NOT GVL_POINT_MANAGER.PointManager.Diag.xZLimitValid THEN
		uiPointCheckReason := UINT#13;
	ELSIF NOT ((stPointCheckCandidate.X >= alrRobotSoftwareMinPosition[1])
		AND (stPointCheckCandidate.X <= alrRobotSoftwareMaxPosition[1])
		AND (stPointCheckCandidate.Y >= alrRobotSoftwareMinPosition[2])
		AND (stPointCheckCandidate.Y <= alrRobotSoftwareMaxPosition[2])
		AND (stPointCheckCandidate.Z >= alrRobotSoftwareMinPosition[3])
		AND (stPointCheckCandidate.Z <= alrRobotSoftwareMaxPosition[3])) THEN
		uiPointCheckReason := UINT#14;
	ELSIF NOT (((stPointCheckCandidate.SpeedFactor > 0.1)
		OR ((uiPointCheckLoop >= UINT#13) AND (stPointCheckCandidate.SpeedFactor >= 0.1)))
		AND (stPointCheckCandidate.SpeedFactor <= 1.0)) THEN
		uiPointCheckReason := UINT#15;
	ELSIF NOT stPointCheckCandidate.xConfigured THEN
		uiPointCheckReason := UINT#16;
	ELSIF NOT xDrivesReady THEN
		uiPointCheckReason := UINT#17;
	ELSIF NOT xPointCheckConnectionAlive THEN
		uiPointCheckReason := UINT#19;
	ELSIF xHmiRobotActionAttempt OR GVL_CELL_CONTROL.xStart OR GVL_CELL_CONTROL.xStop
	OR GVL_CELL_CONTROL.xDisable OR GVL_HMI.xRobotStop OR GVL_HMI.xRobotReset
	OR stSelectedMagazineCommand.xExecute OR stSelectedMagazineCommand.xStop
	OR GVL_CELL_MANAGER.Command.stRobot.xExecute OR GVL_CELL_MANAGER.Command.stRobot.xStop
	OR GVL_MACHINE.Command[1].stRobot.xExecute OR GVL_MACHINE.Command[1].stRobot.xStop
	OR GVL_MACHINE.Command[2].stRobot.xExecute OR GVL_MACHINE.Command[2].stRobot.xStop
	OR GVL_MACHINE.Command[3].stRobot.xExecute OR GVL_MACHINE.Command[3].stRobot.xStop THEN
		uiPointCheckReason := UINT#20;
	END_IF;
	IF (uiPointCheckReason = UINT#0) AND (uiPointCheckMachine > UINT#0) THEN
		IF NOT GVL_MACHINE.Status[uiPointCheckMachine].stIo.xDoorOpen
		OR GVL_MACHINE.Status[uiPointCheckMachine].stIo.xDoorClosed THEN
			uiPointCheckReason := UINT#18;
		END_IF;
	END_IF;
	GVL_HMI.auiPointCheckRejectReason[uiPointCheckLoop] := uiPointCheckReason;
	GVL_HMI.axPointCheckAllowed[uiPointCheckLoop] := uiPointCheckReason = UINT#0;
END_FOR;

IF xPointCheckRequest THEN
	IF GVL_HMI.axPointCheckAllowed[GVL_HMI.uiPointEditorIndex] THEN
		xPointCheckActive := TRUE;
		xPointCheckStopping := FALSE;
		xPointCheckSeenBusy := FALSE;
		xPointCheckSeenDone := FALSE;
		ePointCheckName := ePointEditorName;
		rPointCheckLatchedSpeed := GVL_CELL_SETTINGS.rPointCheckSpeedPercent;
		GVL_HMI.uiPointCheckIndex := GVL_HMI.uiPointEditorIndex;
		GVL_HMI.udiPointCheckRunSeq := GVL_HMI.udiPointEditorCommandSeq;
		GVL_HMI.uiPointCheckState := UINT#1;
		stRobotHmiCommand.eAction := E_ROBOT_ACTION.MOVE_TO_POINT;
		stRobotHmiCommand.eSetPoint := ePointCheckName;
		stRobotHmiCommand.xExecute := TRUE;
		GVL_HMI.stPointEditorResultPoint := GVL_POINT.Points[ePointCheckName];
		GVL_HMI.uiPointEditorResult := UINT#1;
	ELSE
		GVL_HMI.uiPointEditorRejectReason := GVL_HMI.auiPointCheckRejectReason[GVL_HMI.uiPointEditorIndex];
		uiRobotInterfaceWarningCode := WRN_POINT_CHECK_REJECTED;
	END_IF;
	GVL_HMI.udiPointEditorAckSeq := GVL_HMI.udiPointEditorCommandSeq;
END_IF;

// Потеря разрешений во время проверки требует останова, а не только запрета
// следующего старта. Торможение сохраняет обычные инженерные Deceleration/Jerk.
IF xPointCheckActive THEN
	uiPointCheckMachine := UINT#0;
	IF (GVL_HMI.uiPointCheckIndex <= UINT#9) AND ((GVL_HMI.uiPointCheckIndex MOD UINT#3) <> UINT#1) THEN
		uiPointCheckMachine := (GVL_HMI.uiPointCheckIndex - UINT#1) / UINT#3 + UINT#1;
	END_IF;
	IF NOT xPointCheckConnectionAlive OR NOT xHmiConnectionAlive
	OR NOT GVL_CELL_CONTROL.xManual OR GVL_CELL_CONTROL.xGlobalError
	OR GVL_CELL_MANAGER.Status.xRunning OR GVL_HMI.xModbusMode
	OR stSelectedMagazineCommand.xExecute OR stSelectedMagazineCommand.xStop
	OR GVL_CELL_MANAGER.Command.stRobot.xExecute OR GVL_CELL_MANAGER.Command.stRobot.xStop
	OR GVL_MACHINE.Command[1].stRobot.xExecute OR GVL_MACHINE.Command[1].stRobot.xStop
	OR GVL_MACHINE.Command[2].stRobot.xExecute OR GVL_MACHINE.Command[2].stRobot.xStop
	OR GVL_MACHINE.Command[3].stRobot.xExecute OR GVL_MACHINE.Command[3].stRobot.xStop THEN
		xPointCheckStopRequest := TRUE;
	END_IF;
	IF uiPointCheckMachine > UINT#0 THEN
		IF NOT GVL_MACHINE.Status[uiPointCheckMachine].stIo.xDoorOpen
		OR GVL_MACHINE.Status[uiPointCheckMachine].stIo.xDoorClosed THEN
			xPointCheckStopRequest := TRUE;
		END_IF;
	END_IF;
	IF xPointCheckStopRequest AND NOT xPointCheckStopping THEN
		uiRobotInterfaceWarningCode := WRN_POINT_CHECK_INTERRUPTED;
	END_IF;
	xPointCheckStopping := xPointCheckStopping OR xPointCheckStopRequest
		OR GVL_HMI.xRobotStop OR GVL_CELL_CONTROL.xStop OR GVL_CELL_CONTROL.xDisable;
	IF xPointCheckStopping THEN
		stRobotHmiCommand.xExecute := FALSE;
		stRobotHmiCommand.xStop := TRUE;
		xHmiStopAccepted := TRUE;
	END_IF;
END_IF;

ROBOT(
	xUsePhysicalGripperFeedback := GVL_CELL_SETTINGS.eTestEnvironment = E_CELL_TEST_ENVIRONMENT.NORMAL,
	xPhysicalGripperIoReady := GVL_PHYSICAL_IO.xNormalActive,
	stPhysicalGripperFeedback := GVL_PHYSICAL_IO.stGripperFeedback,
	tPhysicalGripperActionTimeout := GVL_CELL_SETTINGS.stMachineTimeouts.tRobotAction,
	axMagazineExchangeInProgress := axTwinMagazineExchangeInProgress,
	xTestInitialize := xTestInitializePulse,
	auiTestGripperContent := GVL_HMI.stTestScenario.auiGripperContent,
	auiTestGripperType := GVL_HMI.stTestScenario.auiGripperType,
	uiTestOrientation := GVL_HMI.stTestScenario.uiOrientation,
	xExternalCommandInhibit := GVL_HMI.xIoEmergencyStopActive,
	stMachine_1_command := GVL_MACHINE.Command[1].stRobot,
	stMachine_2_command := GVL_MACHINE.Command[2].stRobot,
	stMachine_3_command := GVL_MACHINE.Command[3].stRobot,
	stMagazineCommand := stSelectedMagazineCommand,
	stCellCommand := GVL_CELL_MANAGER.Command.stRobot,
	uiBlankPayloadType := GVL_CELL_MANAGER.Command.uiBlankPayloadType,
	uiDetailPayloadType := GVL_CELL_MANAGER.Command.uiDetailPayloadType,
	stHmiCommand := stRobotHmiCommand,
	xReset := GVL_CELL_CONTROL.xReset OR GVL_HMI.xRobotReset,
	xManual := GVL_CELL_CONTROL.xManual AND NOT GVL_CELL_MANAGER.Status.xRunning,
	xMode := GVL_HMI.xModbusMode,
	xGlobalError := GVL_CELL_CONTROL.xGlobalError,
	xEquipmentStopRequired := GVL_MACHINE.Status[1].xCriticalError
		OR GVL_MACHINE.Status[2].xCriticalError
		OR GVL_MACHINE.Status[3].xCriticalError
		OR GVL_MAGAZINE.astStatus[1].xRobotStopRequired
		OR GVL_MAGAZINE.astStatus[2].xRobotStopRequired
		OR (GVL_GEOMETRY_CONTROL.xSupported AND (GVL_GEOMETRY_CONTROL.astStatus[1].xRobotStopRequired
			OR GVL_GEOMETRY_CONTROL.astStatus[2].xRobotStopRequired)),
	xManualRecoveryAllowed := xManualRecoveryActive,
	xModbusBusy := GVL_ROBOT.xModbusBusy,
	xModbusDone := GVL_ROBOT.xModbusDone,
	xModbusError := GVL_ROBOT.xModbusError,
	stModbusStatus := GVL_ROBOT_MODBUS.Status,
	xHmiDrivesEnable := GVL_HMI.xRobotDrivesEnable,
	xHmiDrivesDisable := GVL_HMI.xRobotDrivesDisable,
	xHmiStop := GVL_HMI.xRobotStop,
	xHmiDrivesEnableAccepted := xHmiDrivesEnableAccepted,
	xHmiDrivesDisableAccepted := xHmiDrivesDisableAccepted,
	xHmiStopAccepted := xHmiStopAccepted OR xIoManualActive OR GVL_HMI.xIoEmergencyStopActive,
	xHmiDrivesEnableAllowed := GVL_HMI.stRobotHmiStatus.xDrivesEnableAllowed,
	xHmiDrivesDisableAllowed := GVL_HMI.stRobotHmiStatus.xDrivesDisableAllowed,
	xHmiStopAllowed := GVL_HMI.stRobotHmiStatus.xStopAllowed,
	xHmiPermit := xRobotHmiPermit AND xHmiConnectionAlive,
	xDrivesPowered := xDrivesPowered,
	xDrivesOff := xDrivesOff,
	xDrivesReady := xDrivesReady,
	xDriveError := xDriveError,
	xMotionBusy := xMotionBusy,
	xMotionResetBusy := xMotionResetBusy,
	tSoftMotionResetTimeout := GVL_CELL_SETTINGS.stAxisGroupTimeouts.tGroupTimeout * UINT#2
		+ GVL_CELL_SETTINGS.stAxisTimeouts.tResetTimeout + T#2S,
	xSingleAxisMotionBusy := uiManualAxisOwner > UINT#0,
	xPointCheckActive := xPointCheckActive,
	xTestAbort := xTestAbortActive OR xIoManualActive,
	rPointCheckSpeedPercent := rPointCheckLatchedSpeed,
	lrGroupAccelerationFactor := REAL_TO_LREAL(MIN(
		GVL_CELL_SETTINGS.rRobotAccelerationPercent,
		GVL_CELL_SETTINGS.rRobotDecelerationPercent)) / 100.0,
	lrGroupJerkFactor := REAL_TO_LREAL(GVL_CELL_SETTINGS.rRobotJerkPercent) / 100.0,
	tModbusStartTimeout := GVL_ROBOT_MODBUS_RETAIN.tCommandStartTimeout,
	xSimulationAccelerationEnable := GVL_CELL_SETTINGS.xSimulationAccelerationActive,
	uiSimulationTimeFactor := GVL_CELL_SETTINGS.uiSimulationTimeFactorApplied,
	FaultRequest := stRobotFaultRequest,
	tGripper1OpenTime := GVL_HMI.tGripper1OpenTime,
	tGripper1CloseTime := GVL_HMI.tGripper1CloseTime,
	tGripper2OpenTime := GVL_HMI.tGripper2OpenTime,
	tGripper2CloseTime := GVL_HMI.tGripper2CloseTime,
	tGripperChangeTime := GVL_HMI.tGripperChangeTime,
	stPoint := GVL_POINT.Points,
	stMotionManager := GVL_MOTION_MANAGER.stMotionManager,
	GroupData := GVL_AXIS_GROUP.AxisGroup,
	stPointManager := GVL_POINT_MANAGER.PointManager,
	Command => GVL_ROBOT.Command,
	ModbusCommand => GVL_ROBOT.ModbusCommand,
	Status => GVL_ROBOT.Status,
	Diag => GVL_ROBOT.Diag,
	Error => GVL_ROBOT.Error,
	GripperCommand => GVL_PHYSICAL_IO.stGripperCommand,
	GripperDiag => GVL_ROBOT.GripperDiag,
	GripperError => GVL_ROBOT.GripperError
);

// Проверка держит свою скорость до фактического окончания/останова движения.
tonPointCheckStart(
	IN := xPointCheckActive AND NOT xPointCheckSeenBusy,
	PT := GVL_CELL_SETTINGS.tPointCheckStartTimeout
);
IF xPointCheckActive THEN
	xPointCheckSeenBusy := xPointCheckSeenBusy OR GVL_ROBOT.Status.xBusy;
	// HMI передаёт Execute импульсом. FB_ROBOT в DONE при снятом Execute
	// сбрасывает свой xDone в том же вызове. Motion сохраняет терминальный
	// ответ; запоминаем его только для уже начатой проверки нужной точки.
	xPointCheckSeenDone := xPointCheckSeenDone OR (xPointCheckSeenBusy
		AND GVL_MOTION_MANAGER.stMotionManager.Status.xDone
		AND (GVL_MOTION_MANAGER.stMotionManager.Status.eCurrentPoint = ePointCheckName));
	IF GVL_ROBOT.Status.xError OR tonPointCheckStart.Q THEN
		GVL_HMI.uiPointCheckState := UINT#4;
		xPointCheckStopping := TRUE;
	END_IF;
	IF xPointCheckStopping THEN
		IF NOT GVL_ROBOT.Status.xBusy AND NOT xMotionBusy
		AND NOT GVL_MOTION_MANAGER.stMotionManager.Status.xBusy THEN
			xPointCheckActive := FALSE;
			IF GVL_HMI.uiPointCheckState <> UINT#4 THEN
				GVL_HMI.uiPointCheckState := UINT#3;
			END_IF;
		END_IF;
	ELSIF xPointCheckSeenDone AND NOT GVL_ROBOT.Status.xBusy AND NOT xMotionBusy
	AND NOT GVL_MOTION_MANAGER.stMotionManager.Status.xBusy THEN
		GVL_HMI.uiPointCheckState := UINT#2;
		xPointCheckActive := FALSE;
	END_IF;
END_IF;
// xPointCheckStopping belongs only to the active verification transaction.
// Leaving it latched would make RunMotion stop an unrelated later group move.
IF NOT xPointCheckActive THEN
	xPointCheckStopping := FALSE;
END_IF;

// Команда автоматики запоминается до следующего вызова RunMotion, который
// является единственным владельцем MC_GroupStop и FB_AXIS Stop.
xRobotProgramStopRequest := GVL_ROBOT.Command.xStop AND NOT xHmiStopAccepted;

// В скане запроса xAllowed учитывает его цель, включая безопасность люка.
// Последняя отклонённая цель не должна блокировать следующую попытку HMI.
xHmiRobotStatusPointTargetAllowed := TRUE;
CASE eHmiRobotStatusPoint OF
	E_POINT_NAME.MACHINE_1_INSIDE,
	E_POINT_NAME.MACHINE_1_CHUCK_APROACH,
	E_POINT_NAME.MACHINE_1_CHUCK_POSITION:
		xHmiRobotStatusPointTargetAllowed := GVL_MACHINE.Status[1].stIo.xDoorOpen
			AND NOT GVL_MACHINE.Status[1].stIo.xDoorClosed;
	E_POINT_NAME.MACHINE_2_INSIDE,
	E_POINT_NAME.MACHINE_2_CHUCK_APROACH,
	E_POINT_NAME.MACHINE_2_CHUCK_POSITION:
		xHmiRobotStatusPointTargetAllowed := GVL_MACHINE.Status[2].stIo.xDoorOpen
			AND NOT GVL_MACHINE.Status[2].stIo.xDoorClosed;
	E_POINT_NAME.MACHINE_3_INSIDE,
	E_POINT_NAME.MACHINE_3_CHUCK_APROACH,
	E_POINT_NAME.MACHINE_3_CHUCK_POSITION:
		xHmiRobotStatusPointTargetAllowed := GVL_MACHINE.Status[3].stIo.xDoorOpen
			AND NOT GVL_MACHINE.Status[3].stIo.xDoorClosed;
END_CASE;
xHmiRobotStatusPointAllowed := xHmiRobotActionBaseAllowed
	AND (eHmiRobotStatusAction = E_ROBOT_ACTION.MOVE_TO_POINT)
	AND (eHmiRobotStatusPoint <> E_POINT_NAME.NONE)
	AND xHmiRobotStatusPointTargetAllowed
	AND (
		((eHmiRobotStatusPoint <> E_POINT_NAME.MAGAZINE_SAFE)
		AND (eHmiRobotStatusPoint <> E_POINT_NAME.MAGAZINE_CHANGE)
		AND (eHmiRobotStatusPoint <> E_POINT_NAME.MAGAZINE_IN_SLOT))
		OR (
			(GVL_HMI.uiRobotManualSlot >= UINT#1)
			AND (GVL_HMI.uiRobotManualSlot <= (GVL_CELL_SETTINGS.MagazineRows * GVL_CELL_SETTINGS.MagazineColumns))
			AND (GVL_HMI.uiRobotManualMagazine >= UINT#1)
			AND (GVL_HMI.uiRobotManualMagazine <= UINT#2)
		)
	);
IF xHmiRobotActionAttempt AND (eHmiRobotStatusAction = E_ROBOT_ACTION.MOVE_TO_POINT) THEN
	GVL_HMI.stRobotHmiStatus.xPointsAllowed := xHmiRobotStatusPointAllowed;
ELSE
	// После обработки запроса возвращаем общую готовность. Буфер последней
	// команды остаётся прежним и не отражает выбор новой точки в интерфейсе.
	GVL_HMI.stRobotHmiStatus.xPointsAllowed := xHmiRobotActionBaseAllowed;
END_IF;
GVL_HMI.stRobotHmiStatus.xGripperAllowed := xHmiGripperActionBaseAllowed;
GVL_HMI.stRobotHmiStatus.xGripper1OpenAllowed := xHmiGripperActionBaseAllowed
	AND NOT GVL_ROBOT.Status.xGripper1Open;
GVL_HMI.stRobotHmiStatus.xGripper1CloseAllowed := xHmiGripperActionBaseAllowed
	AND NOT GVL_ROBOT.Status.xGripper1Closed;
GVL_HMI.stRobotHmiStatus.xGripper2OpenAllowed := xHmiGripperActionBaseAllowed
	AND NOT GVL_ROBOT.Status.xGripper2Open;
GVL_HMI.stRobotHmiStatus.xGripper2CloseAllowed := xHmiGripperActionBaseAllowed
	AND NOT GVL_ROBOT.Status.xGripper2Closed;
GVL_HMI.stRobotHmiStatus.xRotateToBlankAllowed := xHmiGripperActionBaseAllowed
	AND NOT GVL_ROBOT.Status.xRotatedToBlank;
GVL_HMI.stRobotHmiStatus.xRotateToDetailAllowed := xHmiGripperActionBaseAllowed
	AND NOT GVL_ROBOT.Status.xRotatedToDetail;
GVL_HMI.stRobotHmiStatus.xCommandBusy := GVL_ROBOT.Status.xBusy
	OR ((GVL_ROBOT.Diag.eState <> E_ROBOT_STATE.IDLE)
		AND (GVL_ROBOT.Diag.eState <> E_ROBOT_STATE.ERROR))
	OR (GVL_ROBOT.GripperDiag.eState = E_GRIPPER_STATE.EXECUTE);
GVL_HMI.stRobotHmiStatus.uiActiveAction := TO_UINT(GVL_ROBOT.Diag.eActiveAction);
GVL_HMI.stRobotHmiStatus.uiActivePoint := TO_UINT(GVL_ROBOT.Diag.eActivePoint);

IF NOT xHmiConnectionAlive THEN
	GVL_HMI.stRobotHmiStatus.eRejectReason := E_HMI_MANUAL_REJECT.HMI_OFFLINE;
ELSIF NOT xRobotHmiPermit THEN
	GVL_HMI.stRobotHmiStatus.eRejectReason := E_HMI_MANUAL_REJECT.MANUAL_MODE_REQUIRED;
ELSIF GVL_HMI.xModbusMode AND NOT GVL_ROBOT_MODBUS.Status.xReady THEN
	GVL_HMI.stRobotHmiStatus.eRejectReason := E_HMI_MANUAL_REJECT.EXTERNAL_ROBOT_NOT_READY;
ELSIF NOT GVL_HMI.xModbusMode AND GVL_CELL_CONTROL.xGlobalError THEN
	GVL_HMI.stRobotHmiStatus.eRejectReason := E_HMI_MANUAL_REJECT.GLOBAL_ERROR_JOG_ONLY;
ELSIF NOT GVL_HMI.xModbusMode AND xDriveError THEN
	GVL_HMI.stRobotHmiStatus.eRejectReason := E_HMI_MANUAL_REJECT.DRIVE_ERROR;
ELSIF NOT GVL_HMI.xModbusMode AND NOT xDrivesPowered THEN
	GVL_HMI.stRobotHmiStatus.eRejectReason := E_HMI_MANUAL_REJECT.DRIVES_DISABLED;
ELSIF GVL_ROBOT.Status.xBusy
	OR ((GVL_ROBOT.Diag.eState <> E_ROBOT_STATE.IDLE)
		AND (GVL_ROBOT.Diag.eState <> E_ROBOT_STATE.ERROR)) THEN
	GVL_HMI.stRobotHmiStatus.eRejectReason := E_HMI_MANUAL_REJECT.ROBOT_BUSY;
ELSIF xHmiRobotActionAttempt AND (eHmiRobotStatusAction = E_ROBOT_ACTION.MOVE_TO_POINT)
	AND NOT xHmiRobotStatusPointTargetAllowed THEN
	GVL_HMI.stRobotHmiStatus.eRejectReason := E_HMI_MANUAL_REJECT.HATCH_CLOSED;
ELSIF NOT GVL_HMI.xModbusMode AND xMotionBusy THEN
	GVL_HMI.stRobotHmiStatus.eRejectReason := E_HMI_MANUAL_REJECT.AXIS_BUSY;
ELSIF NOT GVL_HMI.xModbusMode AND NOT xHmiRobotActionBaseAllowed THEN
	GVL_HMI.stRobotHmiStatus.eRejectReason := E_HMI_MANUAL_REJECT.MOTION_NOT_READY;
ELSE
	GVL_HMI.stRobotHmiStatus.eRejectReason := E_HMI_MANUAL_REJECT.NONE;
END_IF;

IF rtHmiRobotAction.Q AND NOT xHmiRobotActionAllowed THEN
	GVL_ROBOT.Diag.stWarning.uiCode := WRN_HMI_MANUAL_REJECTED;
	GVL_ROBOT.Diag.stWarning.udiSequence := GVL_ROBOT.Diag.stWarning.udiSequence + UDINT#1;
	IF GVL_ROBOT.Diag.stWarning.udiSequence = UDINT#0 THEN
		GVL_ROBOT.Diag.stWarning.udiSequence := UDINT#1;
	END_IF;
END_IF;

IF uiRobotInterfaceWarningCode <> UINT#0 THEN
	GVL_ROBOT.Diag.stWarning.uiCode := uiRobotInterfaceWarningCode;
	GVL_ROBOT.Diag.stWarning.udiSequence := GVL_ROBOT.Diag.stWarning.udiSequence + UDINT#1;
	IF GVL_ROBOT.Diag.stWarning.udiSequence = UDINT#0 THEN
		GVL_ROBOT.Diag.stWarning.udiSequence := UDINT#1;
	END_IF;
	uiRobotInterfaceWarningCode := UINT#0;
END_IF;
END_METHOD

METHOD PRIVATE RunTwoPallet
GVL_TWO_PALLET.xModeChanged := FALSE;
IF NOT xTwinSimulationInitialized THEN
	FOR uiTwin := 1 TO 2 DO
		// Числа используются только для виртуальных SoftMotion-осей.
		GVL_TWO_PALLET.astSimulationConfig[uiTwin].xConfigured := TRUE;
		GVL_TWO_PALLET.astSimulationConfig[uiTwin].xP1LockOut := TRUE;
		GVL_TWO_PALLET.axSimulationAutoSwapEnabled[uiTwin] := TRUE;
		GVL_TWO_PALLET.astSimulationConfig[uiTwin].lrExchange := 0.0;
		GVL_TWO_PALLET.astSimulationConfig[uiTwin].lrWorkP1 := 100.0;
		GVL_TWO_PALLET.astSimulationConfig[uiTwin].lrWorkP2 := 200.0;
		GVL_TWO_PALLET.astSimulationConfig[uiTwin].lrHome := 0.0;
		GVL_TWO_PALLET.astSimulationConfig[uiTwin].lrTolerance := 1.0;
		GVL_TWO_PALLET.astSimulationConfig[uiTwin].lrVelocity := 100.0;
		GVL_TWO_PALLET.astSimulationConfig[uiTwin].lrAcceleration := 200.0;
		GVL_TWO_PALLET.astSimulationConfig[uiTwin].lrDeceleration := 200.0;
		GVL_TWO_PALLET.astSimulationConfig[uiTwin].lrJerk := 1000.0;
		GVL_TWO_PALLET.astSimulationConfig[uiTwin].tCylinder := T#3S;
		GVL_TWO_PALLET.astSimulationConfig[uiTwin].tMove := T#20S;
		GVL_TWO_PALLET.astSimulationConfig[uiTwin].tHome := T#10S;
		GVL_TWO_PALLET.astSimulationConfig[uiTwin].tPulse := T#150MS;
	END_FOR;
	IF NOT GVL_TWO_PALLET.xAutoSwapDefaultsApplied THEN
		FOR uiTwin := 1 TO 2 DO
			GVL_TWO_PALLET.axAutoSwapEnabled[uiTwin] := TRUE;
		END_FOR;
		GVL_TWO_PALLET.xAutoSwapDefaultsApplied := TRUE;
	END_IF;
	xTwinSimulationInitialized := TRUE;
END_IF;
FOR uiTwin := 1 TO 2 DO
	GVL_TWO_PALLET.auiCommand[uiTwin] := UINT#0;
	axMagazineInventoryChanged[uiTwin] := FALSE;
END_FOR;
IF NOT xTwinStartup THEN
	IF GVL_TWO_PALLET.uiMode = 0 THEN
		GVL_HMI.MagazinePitchX := GVL_TWO_PALLET.lrStaticPitchX;
		GVL_HMI.MagazinePitchY := GVL_TWO_PALLET.lrStaticPitchY;
	ELSE
		GVL_HMI.MagazinePitchX := GVL_TWO_PALLET.lrTwinPitchX;
		GVL_HMI.MagazinePitchY := GVL_TWO_PALLET.lrTwinPitchY;
	END_IF;
	FOR uiTwin := 1 TO 2 DO
		// После перезапуска содержимое сохранено, готовность загрузки подтверждается заново.
		GVL_TWO_PALLET.astStore[uiTwin].axLoaded[1] := FALSE;
		GVL_TWO_PALLET.astStore[uiTwin].axLoaded[2] := FALSE;
		IF GVL_TWO_PALLET.uiMode = 0 THEN
			GVL_DETAIL.astMagazine[uiTwin] := GVL_TWO_PALLET.astStatic[uiTwin];
		END_IF;
	END_FOR;
	xTwinStartup := TRUE;
END_IF;
GVL_TWO_PALLET.xModeChangeAllowed := GVL_CELL_CONTROL.xManual
	AND NOT GVL_CELL_MANAGER.Status.xRunning AND NOT GVL_ROBOT.Status.xBusy AND NOT xMotionBusy
	AND xHmiConnectionAlive AND NOT GVL_HMI.xTestSessionActive AND NOT GVL_ROBOT.Status.xBlankAvailable AND NOT GVL_ROBOT.Status.xDetailAvailable
	AND (GVL_ROBOT.Status.uiMagazineContext = 0)
	AND NOT GVL_MAGAZINE.astStatus[1].xEnabled AND NOT GVL_MAGAZINE.astStatus[2].xEnabled
	AND NOT GVL_MAGAZINE.astStatus[1].xBusy AND NOT GVL_MAGAZINE.astStatus[2].xBusy
	AND NOT GVL_TWO_PALLET.astStatus[1].xBusy AND NOT GVL_TWO_PALLET.astStatus[2].xBusy
	AND NOT GVL_TWO_PALLET.astInput[1].xPowered AND NOT GVL_TWO_PALLET.astInput[2].xPowered
	AND NOT GVL_TWO_PALLET.astStatus[1].xError AND NOT GVL_TWO_PALLET.astStatus[2].xError;

udiTwinSnapshot := GVL_HMI.udiTwinCommandSeq;
uiTwinRequestResult := 0;
xTwinInventoryCommand := FALSE;
IF (udiTwinSnapshot <> 0) AND (udiTwinSnapshot <> GVL_HMI.udiTwinAckSeq) THEN
	stTwinRequest := GVL_HMI.stTwinRequest;
	uiTwinRequestResult := 2; // Условие команды не выполнено
	IF (GVL_HMI.udiHmiCommandClockMs - GVL_HMI.udiTwinIssuedAtMs) > 2000 THEN
		uiTwinRequestResult := 4;
	ELSIF (stTwinRequest.uiMagazine = 0) AND (stTwinRequest.uiCommand = 25) THEN
		IF GVL_TWO_PALLET.xModeChangeAllowed AND (stTwinRequest.uiValue <= 1) AND xHmiConnectionAlive THEN
			IF GVL_TWO_PALLET.uiMode <> stTwinRequest.uiValue THEN
				IF GVL_TWO_PALLET.uiMode = 0 THEN
					GVL_TWO_PALLET.lrStaticPitchX := GVL_HMI.MagazinePitchX;
					GVL_TWO_PALLET.lrStaticPitchY := GVL_HMI.MagazinePitchY;
				ELSE
					GVL_TWO_PALLET.lrTwinPitchX := GVL_HMI.MagazinePitchX;
					GVL_TWO_PALLET.lrTwinPitchY := GVL_HMI.MagazinePitchY;
				END_IF;
				GVL_TWO_PALLET.uiMode := stTwinRequest.uiValue;
				GVL_TWO_PALLET.xModeChanged := TRUE;
				FOR uiTwin := 1 TO 2 DO
					axMagazineInventoryChanged[uiTwin] := TRUE;
					IF GVL_TWO_PALLET.uiMode = 0 THEN GVL_DETAIL.astMagazine[uiTwin] := GVL_TWO_PALLET.astStatic[uiTwin]; END_IF;
					// Базы меняются вместе с механикой: старые координаты нельзя молча использовать.
					GVL_POINT.astRetainPoints[13 + uiTwin].xConfigured := FALSE;
					axMagazinePointsReady[uiTwin] := FALSE;
				END_FOR;
				GVL_POINT.Points[E_POINT_NAME.MAGAZINE_1_DETAIL].xConfigured := FALSE;
				GVL_POINT.Points[E_POINT_NAME.MAGAZINE_2_DETAIL].xConfigured := FALSE;
				IF GVL_TWO_PALLET.uiMode = 0 THEN
					GVL_HMI.MagazinePitchX := GVL_TWO_PALLET.lrStaticPitchX; GVL_HMI.MagazinePitchY := GVL_TWO_PALLET.lrStaticPitchY;
				ELSE
					GVL_HMI.MagazinePitchX := GVL_TWO_PALLET.lrTwinPitchX; GVL_HMI.MagazinePitchY := GVL_TWO_PALLET.lrTwinPitchY;
				END_IF;
				xPointTableReady := FALSE;
			END_IF;
			uiTwinRequestResult := 1;
		END_IF;
	ELSIF (stTwinRequest.uiMagazine >= 1) AND (stTwinRequest.uiMagazine <= 2)
		AND (GVL_TWO_PALLET.uiMode = 1) THEN
		uiTwin := stTwinRequest.uiMagazine;
		IF ((stTwinRequest.uiCommand >= 1) AND (stTwinRequest.uiCommand <= 19))
			OR ((stTwinRequest.uiCommand >= 25) AND (stTwinRequest.uiCommand <= 32)) THEN
			GVL_TWO_PALLET.auiCommand[uiTwin] := stTwinRequest.uiCommand;
			GVL_TWO_PALLET.auiValue[uiTwin] := stTwinRequest.uiValue;
			GVL_TWO_PALLET.audiRevision[uiTwin] := stTwinRequest.udiRevision;
		ELSIF (stTwinRequest.uiCommand >= UINT#20)
			AND (stTwinRequest.uiCommand <= UINT#24) THEN
			xTwinInventoryCommand := TRUE; // Проверить по разрешениям текущего скана ПОСЛЕ вызова FB
		ELSIF stTwinRequest.uiCommand = UINT#33 THEN
			IF (stTwinRequest.uiValue <= UINT#1) AND xHmiConnectionAlive THEN
				IF GVL_CELL_SETTINGS.eTestEnvironment = E_CELL_TEST_ENVIRONMENT.SIMULATION THEN
					GVL_TWO_PALLET.axSimulationAutoSwapEnabled[uiTwin] := stTwinRequest.uiValue = UINT#1;
				ELSE
					GVL_TWO_PALLET.axAutoSwapEnabled[uiTwin] := stTwinRequest.uiValue = UINT#1;
				END_IF;
				uiTwinRequestResult := UINT#1;
			END_IF;
		END_IF;
	END_IF;
END_IF;

FOR uiTwin := 1 TO 2 DO
	GVL_TWO_PALLET.astActiveConfig[uiTwin] := GVL_TWO_PALLET.astConfig[uiTwin];
	IF GVL_CELL_SETTINGS.eTestEnvironment = E_CELL_TEST_ENVIRONMENT.SIMULATION THEN
		GVL_TWO_PALLET.astActiveConfig[uiTwin] := GVL_TWO_PALLET.astSimulationConfig[uiTwin];
		xTwinAutoSwapEnabled := GVL_TWO_PALLET.axSimulationAutoSwapEnabled[uiTwin];
	ELSE
		xTwinAutoSwapEnabled := GVL_TWO_PALLET.axAutoSwapEnabled[uiTwin];
	END_IF;
	// Старые RETAIN-параметры сохраняют прежнюю полярность до первой настройки
	// полных сочетаний. Нормализуем только рабочую копию, без записи в RETAIN.
	IF NOT GVL_TWO_PALLET.astActiveConfig[uiTwin].xSignalPatternsConfigured THEN
		GVL_TWO_PALLET.astActiveConfig[uiTwin].uiP1Signals := UINT#38;
		GVL_TWO_PALLET.astActiveConfig[uiTwin].uiP2Signals := UINT#26;
		IF GVL_TWO_PALLET.astActiveConfig[uiTwin].xP1LockOut THEN
			GVL_TWO_PALLET.astActiveConfig[uiTwin].uiP1Signals := UINT#26;
			GVL_TWO_PALLET.astActiveConfig[uiTwin].uiP2Signals := UINT#38;
		END_IF;
		GVL_TWO_PALLET.astActiveConfig[uiTwin].xSignalPatternsConfigured := TRUE;
	END_IF;
	// Legacy power/reset также проходит владельца механизма и его блокировки.
	IF (GVL_TWO_PALLET.auiCommand[uiTwin] = 0) AND (GVL_TWO_PALLET.uiMode = 1) THEN
		IF GVL_HMI.astMagazineCommand[uiTwin].xEnable THEN GVL_TWO_PALLET.auiCommand[uiTwin] := 1; END_IF;
		IF GVL_HMI.astMagazineCommand[uiTwin].xDisable THEN GVL_TWO_PALLET.auiCommand[uiTwin] := 3; END_IF;
		IF GVL_HMI.astMagazineCommand[uiTwin].xStop THEN GVL_TWO_PALLET.auiCommand[uiTwin] := 15; END_IF;
		IF GVL_HMI.astMagazineCommand[uiTwin].xReset
			OR (GVL_CELL_CONTROL.xReset AND GVL_TWO_PALLET.astStatus[uiTwin].xResetAllowed) THEN
			GVL_TWO_PALLET.auiCommand[uiTwin] := 16;
		END_IF;
	END_IF;

	// Единственное место преобразования транспортных номеров HMI в интерфейс FB.
	astTwinCommand[uiTwin].xEnable := GVL_TWO_PALLET.auiCommand[uiTwin] = UINT#1;
	astTwinCommand[uiTwin].xConfirm := GVL_TWO_PALLET.auiCommand[uiTwin] = UINT#2;
	astTwinCommand[uiTwin].xStart := GVL_TWO_PALLET.auiCommand[uiTwin] = UINT#27;
	astTwinCommand[uiTwin].xRejectStart := GVL_TWO_PALLET.auiCommand[uiTwin] = UINT#28;
	astTwinCommand[uiTwin].xDisable := GVL_TWO_PALLET.auiCommand[uiTwin] = UINT#3;
	astTwinCommand[uiTwin].xSwap := GVL_TWO_PALLET.auiCommand[uiTwin] = UINT#4;
	astTwinCommand[uiTwin].xPowerOn := GVL_TWO_PALLET.auiCommand[uiTwin] = UINT#5;
	astTwinCommand[uiTwin].xPowerOff := GVL_TWO_PALLET.auiCommand[uiTwin] = UINT#6;
	astTwinCommand[uiTwin].xDriveReset := GVL_TWO_PALLET.auiCommand[uiTwin] = UINT#7;
	astTwinCommand[uiTwin].xHome := GVL_TWO_PALLET.auiCommand[uiTwin] = UINT#8;
	astTwinCommand[uiTwin].xLower := GVL_TWO_PALLET.auiCommand[uiTwin] = UINT#9;
	astTwinCommand[uiTwin].xRaise := GVL_TWO_PALLET.auiCommand[uiTwin] = UINT#10;
	astTwinCommand[uiTwin].xSelectPallet := (GVL_TWO_PALLET.auiCommand[uiTwin] = UINT#11)
		OR (GVL_TWO_PALLET.auiCommand[uiTwin] = UINT#12);
	astTwinCommand[uiTwin].xLockIn := GVL_TWO_PALLET.auiCommand[uiTwin] = UINT#29;
	astTwinCommand[uiTwin].xLockOut := GVL_TWO_PALLET.auiCommand[uiTwin] = UINT#30;
	astTwinCommand[uiTwin].xStopIn := GVL_TWO_PALLET.auiCommand[uiTwin] = UINT#31;
	astTwinCommand[uiTwin].xStopOut := GVL_TWO_PALLET.auiCommand[uiTwin] = UINT#32;
	astTwinCommand[uiTwin].xMoveToExchange := GVL_TWO_PALLET.auiCommand[uiTwin] = UINT#13;
	astTwinCommand[uiTwin].xMoveToWork := GVL_TWO_PALLET.auiCommand[uiTwin] = UINT#14;
	astTwinCommand[uiTwin].xStop := GVL_TWO_PALLET.auiCommand[uiTwin] = UINT#15;
	astTwinCommand[uiTwin].xReset := GVL_TWO_PALLET.auiCommand[uiTwin] = UINT#16;
	astTwinCommand[uiTwin].xJogPositive := GVL_TWO_PALLET.auiCommand[uiTwin] = UINT#17;
	astTwinCommand[uiTwin].xJogNegative := GVL_TWO_PALLET.auiCommand[uiTwin] = UINT#18;
	astTwinCommand[uiTwin].xJogRelease := GVL_TWO_PALLET.auiCommand[uiTwin] = UINT#19;
	astTwinCommand[uiTwin].xTeachOperator := GVL_TWO_PALLET.auiCommand[uiTwin] = UINT#25;
	astTwinCommand[uiTwin].xTeachWork := GVL_TWO_PALLET.auiCommand[uiTwin] = UINT#26;
	astTwinCommand[uiTwin].uiPallet := GVL_TWO_PALLET.auiValue[uiTwin];
	IF GVL_TWO_PALLET.auiCommand[uiTwin] = UINT#11 THEN
		astTwinCommand[uiTwin].uiPallet := UINT#1;
	ELSIF GVL_TWO_PALLET.auiCommand[uiTwin] = UINT#12 THEN
		astTwinCommand[uiTwin].uiPallet := UINT#2;
	END_IF;
	astTwinCommand[uiTwin].udiRevision := GVL_TWO_PALLET.audiRevision[uiTwin];

